// TwinCAT 3 PLC project Test
// ProgramVersion: 3.1.4026.26
// CompilerDefines: VISU_USEPROPERTYINFO
// libraries:
//   Tc2_Standard, * (Beckhoff Automation GmbH)
//   Tc2_System, * (Beckhoff Automation GmbH)
//   VisuDialogs, * (System)
//   VisuDialogs
// project tree:
//   DUTs/ Auto_Test_DB_DUT.TcDUT, Auto_Test_DUT.TcDUT, Barcode_Station_DUT.TcDUT, Charger_DUT.TcDUT, Gate_Station_DUT.TcDUT, Level_Keys_DUT.TcDUT, Profiling_Station_DUT.TcDUT, Shuttle_Position_UDT.TcDUT, U_DWORD_REAL1.TcDUT
//   DUTs/Carousel/ Chain_Control_DUT.TcDUT, Chain_Settings_DUT.TcDUT, E_Carousel_PopUpMotor.TcDUT, PopUp_Control_DUT.TcDUT, PopUp_Inputs_DUT.TcDUT, PopUp_Instruction_DUT.TcDUT, PopUp_Motors_DUT.TcDUT, PopUp_Motor_Settings_DUT.TcDUT, PopUp_Settings_DUT.TcDUT, PopUp_Side_Status_DUT.TcDUT, Roller_Control_DUT.TcDUT, Roller_Inputs_DUT.TcDUT, Roller_Instruction_DUT.TcDUT, Roller_Settings_DUT.TcDUT, TBCnv_Control_DUT.TcDUT, TBCnv_Settings_DUT.TcDUT, Turn_Table_Control_DUT.TcDUT, Turn_Table_Inputs_DUT.TcDUT, Turn_Table_Instruction_DUT.TcDUT, Turn_Table_Motor_DUT.TcDUT, Turn_Table_Settings_DUT.TcDUT
//   DUTs/Conveyors/ Buffer_Cnv_Control_DUT.TcDUT, Buffer_Cnv_Inputs_DUT.TcDUT, Buffer_Cnv_Settings_DUT.TcDUT, Cnv_Errors_DUT.TcDUT, Cnv_Inputs_DUT.TcDUT, Cnv_Instruction_DUT.TcDUT, Cnv_Interlock_DUT.TcDUT, Cnv_Level_Control_DUT.TcDUT, Cnv_Level_Inputs_DUT.TcDUT, Cnv_Level_Settings_DUT.TcDUT, Cnv_Motor_DUT.TcDUT, Cnv_Motor_Settings_DUT.TcDUT, Cnv_VTD_Control_DUT.TcDUT, Cnv_VTD_Settings_DUT.TcDUT, ECnv_Control_DUT.TcDUT, ECnv_Settings_DUT.TcDUT
//   DUTs/HMI/ ST_HMI_ConveyorCommand.TcDUT, ST_HMI_ConveyorStatus.TcDUT, ST_HMI_DeviceSummary.TcDUT, ST_HMI_GateCommand.TcDUT, ST_HMI_GateStatus.TcDUT, ST_HMI_GateSummary.TcDUT, ST_HMI_SystemCommand.TcDUT, ST_HMI_SystemStatus.TcDUT, ST_HMI_VtdCommand.TcDUT, ST_HMI_VtdOverview.TcDUT, ST_HMI_VtdStatus.TcDUT, ST_VTD_ManualHmiCommand.TcDUT, ST_VTD_ManualHmiStatus.TcDUT, ST_VTD_ManualSettings.TcDUT, ST_VTD_PdHmiCommand.TcDUT, ST_VTD_PdHmiStatus.TcDUT
//   DUTs/Safety_Stops/ Sfts_Control_DUT.TcDUT, Sfts_Inputs_DUT.TcDUT, Sfts_Instruction_DUT.TcDUT, Sfts_Settings_DUT.TcDUT
//   DUTs/SEW/ E_SEW_MovikitMode.TcDUT, ST_SEW_MovikitStatus.TcDUT, ST_SEW_ProcessInput5.TcDUT, ST_SEW_ProcessInput8.TcDUT, ST_SEW_VelocityScaling.TcDUT, ST_SEW_VelocityStatus.TcDUT
//   DUTs/System/ E_BarcodeState.TcDUT, ID_Decoded_DUT.TcDUT, OrderTable_DUT.TcDUT, System_DUT.TcDUT, System_Settings_DUT.TcDUT, WMS_OPC_UA_DUT.TcDUT
//   DUTs/VTD/ VTD_Control_DUT.TcDUT, VTD_Errors_DUT.TcDUT, VTD_Inputs_DUT.TcDUT, VTD_Instruction_DUT.TcDUT, VTD_Levels_DUT.TcDUT, VTD_Motor_DUT.TcDUT, VTD_Outputs_DUT.TcDUT, VTD_Settings_DUT.TcDUT, VTD_Shuttle_Interlock_DUT.TcDUT
//   / GlobalTextList.TcGTLO, PlcTask.TcTTO, TL_Test.TcTLO, Visualization Manager.TcVMO (not stored), VISU_TASK.TcTTO
//   GVLs/ Control.TcGVL, Errors.TcGVL, Settings.TcGVL, System.TcGVL, System_Control.TcGVL
//   GVLs/HMI/ CNV_HMI.TcGVL, CNV_HMI_IO.TcGVL, GVL_HMI_Carousel.TcGVL, GVL_HMI_CNV.TcGVL, GVL_HMI_Gates.TcGVL, GVL_HMI_System.TcGVL, GVL_HMI_VTD.TcGVL
//   GVLs/IO/ IO_Cards.TcGVL, IO_Chargers.TcGVL, IO_RemoteModules.TcGVL, IO_Safety.TcGVL, IO_VFDs.TcGVL
//   POUs/Conveyors/ Buffer_Conveyor_FB.TcPOU, FB_Conveyor_MotorInterlock.TcPOU
//   POUs/ DWORD_REAL.TcPOU, Inputs.TcPOU, MAIN.TcPOU, Outputs.TcPOU, Profile_Station_FC.TcPOU, Stack_Lights_FB.TcPOU
//   POUs/SEW/ FB_SEW_Drive.TcPOU, FB_SEW_ProcessDataTest.TcPOU, FB_SEW_VelocityDrive.TcPOU, FC_SEW_MovikitModeName.TcPOU, FC_VTD_PdHmiUpdateStatus.TcPOU
//   POUs/System/ Barcode_Station_FB.TcPOU, Conveyors_Transfer.TcPOU
//   POUs/System/Functions/ ByteArrayToString.TcPOU, FC_TIAParseDINT.TcPOU, FC_TIAScalarToken.TcPOU, FindBoolField.TcPOU, FindDINTFieldFragmented.TcPOU, FindIntField.TcPOU, FindINTFieldFragmented.TcPOU, FindStringField.TcPOU, ID_Decode_F.TcPOU, RemovePlusSign.TcPOU, Set_Bit_F.TcPOU
//   POUs/System/Tests/ FC_TestTIAFoundation.TcPOU, FC_TestTIAParsing.TcPOU
//   POUs/VTD/ FB_VTD_ManualControl.TcPOU, Light_Bars_FB.TcPOU, VTD_FB.TcPOU
//   VISUs/ Access_Gates.TcVIS, Alarms.TcVIS, Carrousel.TcVIS, CNV.TcVIS, CNV_Settings.TcVIS, Dialog.TcVIS, FP_Conveyor.TcVIS, FP_Drive.TcVIS, FP_Test.TcVIS, Header.TcVIS, ImagePool.TcIPO (not stored), Main.TcVIS, NavBar.TcVIS, Order_Table.TcVIS, Shuttles.TcVIS, teste.TcVIS, Visualization.TcVIS, VISU_Seeds.TcVIS, VTD.TcVIS, VTDManualTest.TcVIS, VTD_Settings.TcVIS
// real-time tasks:
//   TASK IoTask: cycle T#10ms, priority 1, ADS port 301
//   TASK PlcTask: cycle T#10ms, priority 20, ADS port 350
//   TASK VISU_TASK: cycle T#200000us, priority 30, ADS port 351
// I/O:
//   DEVICE Device 1 (EtherCAT), AmsNetId 10.1.179.234.2.1
//     Term 30 (EK1200) [EK1200-5000 EtherCAT Power supply (2A E-Bus)]
//       Term 3 (EL1809) [EL1809 16Ch. Dig. Input 24V, 3ms]
//       Term 4 (EL1809) [EL1809 16Ch. Dig. Input 24V, 3ms]
//       Term 5 (EL2809) [EL2809 16Ch. Dig. Output 24V, 0.5A]
//       Term 6 (EL2809) [EL2809 16Ch. Dig. Output 24V, 0.5A]
//       Term 7 (EL6910) [EL6910, TwinSAFE PLC]
//       Term 8 (EL1918) [EL1918, 8Ch. Safety Input 24V, TwinSAFE]
//         modules: Module 1 (FSOE), Module 2 (FSLOGIC)
//       Term 9 (EL2912) [EL2912, 2Ch. Safety Output 24V, 2A, TwinSAFE]
//         modules: Module 1 (FSOE), Module 2 (FSOUT), Module 3 (DEVICEIO), Module 4 (FSLOGIC)
//       Term 10 (EL9410) [EL9410 E-Bus Power Supplier  (Diagnostics)]
//       Term 11 (EK1322) [EK1322 2-port EtherCAT P junction with feed-in]
//       Term 12 (EK1322) [EK1322 2-port EtherCAT P junction with feed-in]
//       Term 13 (EK1322) [EK1322 2-port EtherCAT P junction with feed-in]
//         Box 14 (EPP2328-0002) [EPP2328-0002 4 CH. Dig. In, 3ms, 4 Ch. Dig. Out 24V, 2A, M12]
//       Term 43 (EL6633) [EL6633 PROFINET IO Controller]
//       Term 16 (EK1122) [EK1122 2 port EtherCAT junction]
//         Box 17 (CU1124) [CU1124 EtherCAT junction (4-ports)]
//         Box 19 (CU1128) [CU1128 6x EtherCAT junction]
//           Term 22 (CU1128-B) [CU1128 6x EtherCAT junction - Dev A]
//           Term 23 (CU1128-C) [CU1128 6x EtherCAT junction - Dev B]
//             Box 24 (MOVI-C Decentralized Electronics) [MOVI-C Decentralized Electronics]
//               modules: Module 1 (Standard 16 PD), Module 2 (Failsafe Container 28 Byte)
//             Box 25 (MOVI-C Decentralized Electronics) [MOVI-C Decentralized Electronics]
//               modules: Module 1 (Standard 16 PD), Module 2 (FSoE Safety IO 48 bit)
//             Box 45 (MOVI-C Decentralized Electronics) [MOVI-C Decentralized Electronics]
//               modules: Module 1 (Standard 16 PD), Module 2 (Failsafe Container 28 Byte)
//             Box 1 (MOVI-C MOVIPRO) [MOVI-C MOVIPRO]
//               modules: Module 1 (Standard 16 PD), Module 2 (FSoE Safety IO 48 bit)
//             Box 27 (MOVI-C Decentralized Electronics) [MOVI-C Decentralized Electronics]
//               modules: Module 1 (Standard 16 PD)
//             Box 47 (MOVI-C Decentralized Electronics) [MOVI-C Decentralized Electronics]
//               modules: Module 1 (Standard 16 PD)
//             Box 48 (MOVI-C Decentralized Electronics) [MOVI-C Decentralized Electronics]
//               modules: Module 1 (Standard 16 PD)
//             Box 49 (MOVI-C Decentralized Electronics) [MOVI-C Decentralized Electronics]
//               modules: Module 1 (Standard 16 PD)
//             Box 53 (MOVI-C Decentralized Electronics) [MOVI-C Decentralized Electronics]
//               modules: Module 1 (Standard 16 PD)
//   DEVICE Device 4 (COM Port)
// variable links:
//   Device 1 (EtherCAT) <-> Device 1 (EtherCAT)/Term 30 (EK1200)/Term 16 (EK1122)/Box 19 (CU1128)/Term 23 (CU1128-C)/Box 1 (MOVI-C MOVIPRO)
//     Term 30 (EK1200)/Term 7 (EL6910)/ConnectionInputs/Message_14 TxPDO <-> Module 2 (FSoE Safety IO 48 bit)/FSoE Safety Outputs 48 bit/FSOE
//     Term 30 (EK1200)/Term 7 (EL6910)/ConnectionOutputs/Message_14 RxPDO <-> Module 2 (FSoE Safety IO 48 bit)/FSoE Safety Inputs 48 bit/FSOE
//   Device 1 (EtherCAT) <-> Device 1 (EtherCAT)/Term 30 (EK1200)/Term 8 (EL1918)
//     Term 30 (EK1200)/Term 7 (EL6910)/ConnectionInputs/Message_13 TxPDO <-> Module 1 (FSOE)/FSoE Outputs/FSOE
//     Term 30 (EK1200)/Term 7 (EL6910)/ConnectionOutputs/Message_13 RxPDO <-> Module 1 (FSOE)/FSoE Inputs/FSOE
//   Test/Test Instance <-> Device 1 (EtherCAT)/Term 30 (EK1200)/Term 16 (EK1122)/Box 19 (CU1128)/Term 23 (CU1128-C)/Box 1 (MOVI-C MOVIPRO)
//     PlcTask Inputs/IO_VFDs.VTD_EcState <-> InfoData/State
//     PlcTask Inputs/IO_VFDs.VTD_PI_01 <-> Module 1 (Standard 16 PD)/Inputs 16 PD/PI 1
//     PlcTask Inputs/IO_VFDs.VTD_PI_02 <-> Module 1 (Standard 16 PD)/Inputs 16 PD/PI 2
//     PlcTask Inputs/IO_VFDs.VTD_PI_03 <-> Module 1 (Standard 16 PD)/Inputs 16 PD/PI 3
//     PlcTask Inputs/IO_VFDs.VTD_PI_04 <-> Module 1 (Standard 16 PD)/Inputs 16 PD/PI 4
//     PlcTask Inputs/IO_VFDs.VTD_PI_05 <-> Module 1 (Standard 16 PD)/Inputs 16 PD/PI 5
//     PlcTask Inputs/IO_VFDs.VTD_PI_06 <-> Module 1 (Standard 16 PD)/Inputs 16 PD/PI 6
//     PlcTask Inputs/IO_VFDs.VTD_PI_07 <-> Module 1 (Standard 16 PD)/Inputs 16 PD/PI 7
//     PlcTask Inputs/IO_VFDs.VTD_PI_08 <-> Module 1 (Standard 16 PD)/Inputs 16 PD/PI 8
//     PlcTask Inputs/IO_VFDs.VTD_WcState <-> WcState/WcState
//     PlcTask Outputs/IO_VFDs.VTD_PO_01 <-> Module 1 (Standard 16 PD)/Outputs 16 PD/PO 1
//     PlcTask Outputs/IO_VFDs.VTD_PO_02 <-> Module 1 (Standard 16 PD)/Outputs 16 PD/PO 2
//     PlcTask Outputs/IO_VFDs.VTD_PO_03 <-> Module 1 (Standard 16 PD)/Outputs 16 PD/PO 3
//     PlcTask Outputs/IO_VFDs.VTD_PO_04 <-> Module 1 (Standard 16 PD)/Outputs 16 PD/PO 4
//     PlcTask Outputs/IO_VFDs.VTD_PO_05 <-> Module 1 (Standard 16 PD)/Outputs 16 PD/PO 5
//     PlcTask Outputs/IO_VFDs.VTD_PO_06 <-> Module 1 (Standard 16 PD)/Outputs 16 PD/PO 6
//     PlcTask Outputs/IO_VFDs.VTD_PO_07 <-> Module 1 (Standard 16 PD)/Outputs 16 PD/PO 7
//     PlcTask Outputs/IO_VFDs.VTD_PO_08 <-> Module 1 (Standard 16 PD)/Outputs 16 PD/PO 8
//   Test/Test Instance <-> Device 1 (EtherCAT)/Term 30 (EK1200)/Term 7 (EL6910)
//     PlcTask Outputs/IO_Safety.ErrorAcknowledgement <-> StandardOutputs/Standard In Var 1
//     PlcTask Outputs/IO_Safety.Run <-> StandardOutputs/Standard In Var 2
//     PlcTask Outputs/IO_Safety.SEW_Safety_Reset <-> StandardOutputs/Standard In Var 10

CONFIGURATION Test
    RESOURCE PLC ON TwinCAT3
        TASK PlcTask(INTERVAL := T#10ms, PRIORITY := 20);
        TASK VISU_TASK(INTERVAL := T#200000us, PRIORITY := 30);
        PROGRAM MAIN WITH PlcTask : MAIN;
        PROGRAM VisuElems_Visu_Prg WITH VISU_TASK : VisuElems.Visu_Prg;
    END_RESOURCE
END_CONFIGURATION

// ---- DUTs/Auto_Test_DB_DUT.TcDUT
TYPE Auto_Test_DB_DUT :
STRUCT
	System: ARRAY[1..5] OF Auto_Test_DUT;
END_STRUCT
END_TYPE

// ---- DUTs/Auto_Test_DUT.TcDUT
TYPE Auto_Test_DUT :
STRUCT
	Duration:	TIME;
	Start_Time:	STRING[20];
	Stop_Time:	STRING[20];
	Time_Running:	TIME;
	Total_Duration:	TIME;
END_STRUCT
END_TYPE

// ---- DUTs/Barcode_Station_DUT.TcDUT
TYPE Barcode_Station_DUT :
STRUCT
	// Explicit capacity matches the default STRING length in the Siemens source.
	Start:	BOOL;
	Ready:	BOOL;
	Running:	BOOL;
	Done:	BOOL;
	Valid:	BOOL;
	Reading_Gate_number:	STRING(254);
	Reading_Gate_number_OLD:	STRING(254);
	Number_OF_Reading_Gates:	STRING(254);
	Number_OF_Reading_Gates_OLD:	STRING(254);
	Barcode:	STRING(254);
	Barcode_Old:	STRING(254);
END_STRUCT
END_TYPE

// ---- DUTs/Carousel/Chain_Control_DUT.TcDUT
// Internal state of the carousel chain conveyor (Control.Chain_Cnv).
// Same layout as ECnv_Control_DUT. Drive: SEW MOVIKIT Velocity Drive, 5 PD.
TYPE Chain_Control_DUT :
STRUCT
	Mode:	UINT;	// 0 Disabled, 1 Manual, 2 Semi-Auto, 3 Auto, 5 Maintenance
	Error:	BOOL;
	Warning:	UINT;
	Enabled:	BOOL;
	Stopped:	BOOL;
	Done:	BOOL;
	Running:	BOOL;
	Ready_For_Task:	BOOL;
	Current_Task_Type:	UINT;
	Current_Task_ID:	UINT;
	Cnv_Occupied:	BOOL;
	SM_State:	UINT;	// State machine value
	Motor:	Cnv_Motor_DUT;
	Instruction:	Cnv_Instruction_DUT;
	Inputs:	Cnv_Inputs_DUT;	// Forward/Backward_Sensor; VFD_* words not used with SEW
	Cnv_Errors:	Cnv_Errors_DUT;
END_STRUCT
END_TYPE

// ---- DUTs/Carousel/Chain_Settings_DUT.TcDUT
// Parameters of the carousel chain conveyor (Settings.Chain_Cnv). Based on ECnv_Settings_DUT.
// 0 = not configured: the function that uses the value is blocked.
TYPE Chain_Settings_DUT :
STRUCT
	ID:	DINT;	// XXYYZZ
	Motor:	Cnv_Motor_Settings_DUT;	// Same name as Control.<device>.Motor
END_STRUCT
END_TYPE

// ---- DUTs/Carousel/E_Carousel_PopUpMotor.TcDUT
// Motor of a carousel popup that is allowed to run (Control.Pop_Up_Cnv[n].Active_Motor).
// The values are the motor indices of the popup's FB_Conveyor_MotorInterlock instance.
{attribute 'qualified_only'}
TYPE E_Carousel_PopUpMotor :
(
    None := 0,          // No motor granted
    Lift := 1,          // Motors.Lift
    Transfer := 2       // Motors.Transfer
) INT;
END_TYPE

// ---- DUTs/Carousel/PopUp_Control_DUT.TcDUT
// Internal state of one carousel popup (Control.Pop_Up_Cnv[1..2]): lift + transfer conveyor.
// Based on Dallas PopUp_Cnv_Control; same header as ECnv_Control_DUT / Buffer_Cnv_Control_DUT.
// Motors.Lift and Motors.Transfer never run at the same time (Active_Motor, FB_Conveyor_MotorInterlock).
// Drives: SEW MOVIKIT Velocity Drive, 5 PD (Motor.stProcessInput / aProcessOutput in Cnv_Motor_DUT).
TYPE PopUp_Control_DUT :
STRUCT
	Mode:	UINT;	// 0 Disabled, 1 Manual, 2 Semi-Auto, 3 Auto, 5 Maintenance
	Error:	BOOL;
	Warning:	UINT;
	Enabled:	BOOL;
	Stopped:	BOOL;
	Done:	BOOL;
	Running:	BOOL;
	Ready_For_Task:	BOOL;
	Current_Task_Type:	UINT;
	Current_Task_ID:	UINT;
	Cnv_Occupied:	BOOL;
	SM_State:	UINT;	// State machine value
	Active_Side:	INT;	// Side 1..4 of the running transfer, 0 = none
	Inputs:	PopUp_Inputs_DUT;
	Side:	ARRAY[1..4] OF PopUp_Side_Status_DUT;	// 1/2 transfer Fwd/Rev end (Lift_Up), 3/4 Lift_Down level (pallet moved by the neighbour, e.g. Chain_Cnv)

	// Motor group: one motor at a time
	Motors:	PopUp_Motors_DUT;
	Active_Motor:	E_Carousel_PopUpMotor;	// Motor allowed to run, None = no motor granted
	Motor_Changeover:	BOOL;	// A motor is requested and waits until the other one stopped + Changeover_Time

	Instruction:	PopUp_Instruction_DUT;
	Cnv_Errors:	Cnv_Errors_DUT;
END_STRUCT
END_TYPE

// ---- DUTs/Carousel/PopUp_Inputs_DUT.TcDUT
// Sensors of one carousel popup (Control.Pop_Up_Cnv[n].Inputs). Written only by FC Inputs.
// Based on Dallas PopUp_Cnv_Inputs ("Lift Up" / "Lift Down") plus the popup pallet sensor.
// TRUE = condition present (invert NC sensors in FC Inputs).
TYPE PopUp_Inputs_DUT :
STRUCT
	Lift_Up:	BOOL;	// Lift at the top = transfer conveyor level
	Lift_Down:	BOOL;	// Lift at the bottom = chain level (pallet on Chain_Cnv, to confirm with the layout)
	Pallet_Present:	BOOL;	// Pallet on the popup (end of an inbound transfer)
END_STRUCT
END_TYPE

// ---- DUTs/Carousel/PopUp_Instruction_DUT.TcDUT
// Commands of one carousel popup (WMS / order table / HMI). Same members as Dallas PopUp_Cnv_Instruction.
TYPE PopUp_Instruction_DUT :
STRUCT
	Mode_Change:	UINT;	// Requested mode, see Mode
	Stop:	BOOL;
	Enable:	BOOL;
	Reset:	BOOL;
	Execute:	BOOL;	// Rising edge starts the task
	Task_ID:	UINT;
	Task_Metadata:	STRING;
	Transfer_To_ID:	DINT;	// Outbound: ID (XXYYZZ) of the receiving device
	Transfer_From_ID:	DINT;	// Inbound: ID (XXYYZZ) of the sending device
	Transfer_in_Progress:	BOOL;	// Written by the conveyor FB
	Inbound_Ready:	BOOL;	// Written by Conveyors_Transfer
	Transfer_Complete:	BOOL;
	Outbound_Ready:	BOOL;	// Written by Conveyors_Transfer
	Start_Transfer:	BOOL;
	Start_Transfer_Backward:	BOOL;	// Manual mode only

	// Manual mode
	Transfer_Fwd:	BOOL;	// Jog the transfer conveyor forward (only at Lift_Up)
	Transfer_Bwd:	BOOL;	// Jog the transfer conveyor backward (only at Lift_Up)
	Lift_Up:	BOOL;	// Auto: move the lift up. Manual: jog up
	Lift_Down:	BOOL;	// Auto: move the lift down. Manual: jog down
END_STRUCT
END_TYPE

// ---- DUTs/Carousel/PopUp_Motors_DUT.TcDUT
// Motors of one carousel popup (Control.Pop_Up_Cnv[n].Motors). They never run at the same time:
// PopUp_Conveyor_FB grants one motor at a time (FB_Conveyor_MotorInterlock, Active_Motor).
// Drives: SEW MOVIKIT Velocity Drive, 5 PD.
TYPE PopUp_Motors_DUT :
STRUCT
	Lift:	Cnv_Motor_DUT;	// Lift up / down (E_Carousel_PopUpMotor.Lift)
	Transfer:	Cnv_Motor_DUT;	// Transfer conveyor, runs only at Lift_Up (E_Carousel_PopUpMotor.Transfer)
END_STRUCT
END_TYPE

// ---- DUTs/Carousel/PopUp_Motor_Settings_DUT.TcDUT
// Motor parameters of one carousel popup (Settings.Pop_Up_Cnv[n].Motors).
// Same member names as PopUp_Motors_DUT in Control.
TYPE PopUp_Motor_Settings_DUT :
STRUCT
	Lift:	Cnv_Motor_Settings_DUT;	// Transfer_Time = lift travel watchdog
	Transfer:	Cnv_Motor_Settings_DUT;
END_STRUCT
END_TYPE

// ---- DUTs/Carousel/PopUp_Settings_DUT.TcDUT
// Parameters of one carousel popup (Settings.Pop_Up_Cnv[1..2]). Based on Dallas PopUp_Cnv_Settings;
// the G120 hardware IDs are replaced by the SEW scaling of each drive (Motors.<motor>.Drive).
// 0 = not configured: the function that uses the value is blocked.
TYPE PopUp_Settings_DUT :
STRUCT
	ID:	DINT;	// XXYYZZ
	Side_ID:	ARRAY[1..4] OF DINT;	// Neighbour ID per side, 0 = none. 1/2 transfer Fwd/Rev end (Lift_Up), 3/4 Lift_Down level
	Side_Boost_Time:	ARRAY[1..4] OF UINT;	// [s] start boost per side, 0 = none (Dallas TimeStartBoost_PxToPy)
	Boost_Speed:	UINT := 100;	// Units of Motors.Transfer.Speed

	// Motor group: Lift and Transfer never run at the same time
	Motors:	PopUp_Motor_Settings_DUT;
	Changeover_Time:	UINT;	// [ms] all motors stopped before the other motor may start (brake closed), 0 = not configured
END_STRUCT
END_TYPE

// ---- DUTs/Carousel/PopUp_Side_Status_DUT.TcDUT
// Device on one side of a popup (Control.Pop_Up_Cnv[n].Side[1..4]). Written every cycle by Conveyors_Transfer.
// Replaces the hard-coded neighbour reads of the Dallas PConveyor FBs.
TYPE PopUp_Side_Status_DUT :
STRUCT
	In_Position:	BOOL;	// Neighbour aligned with the popup (VTD at the level, turntable at the station). TRUE for fixed conveyors
	Inbound_Ready:	BOOL;	// Neighbour can receive a pallet
	Running:	BOOL;	// Neighbour transport motor turning (handshake before sending)
	Occupied:	BOOL;	// Neighbour detects the pallet (end of an outbound transfer)
END_STRUCT
END_TYPE

// ---- DUTs/Carousel/Roller_Control_DUT.TcDUT
// Internal state of one carousel roller conveyor (Control.Roller_Cnv[1..5]).
// Same layout as ECnv_Control_DUT. Drive: SEW MOVIKIT Velocity Drive, 5 PD.
TYPE Roller_Control_DUT :
STRUCT
	Mode:	UINT;	// 0 Disabled, 1 Manual, 2 Semi-Auto, 3 Auto, 5 Maintenance
	Error:	BOOL;
	Warning:	UINT;
	Enabled:	BOOL;
	Stopped:	BOOL;
	Done:	BOOL;
	Running:	BOOL;
	Ready_For_Task:	BOOL;
	Current_Task_Type:	UINT;
	Current_Task_ID:	UINT;
	Cnv_Occupied:	BOOL;
	SM_State:	UINT;	// State machine value
	Motor:	Cnv_Motor_DUT;
	Instruction:	Roller_Instruction_DUT;
	Inputs:	Roller_Inputs_DUT;
	Cnv_Errors:	Cnv_Errors_DUT;
END_STRUCT
END_TYPE

// ---- DUTs/Carousel/Roller_Inputs_DUT.TcDUT
// Sensors of one carousel roller conveyor (Control.Roller_Cnv[n].Inputs). Written only by FC Inputs.
// Based on Cnv_Inputs_DUT and Dallas Inbound/Outbound_Cnv_Inputs. The VFD_* words are not needed:
// with SEW the drive data is in Motor.stProcessInput. TRUE = condition present (invert NC sensors in FC Inputs).
TYPE Roller_Inputs_DUT :
STRUCT
	Forward_Sensor:	BOOL;	// Pallet at the forward end
	Backward_Sensor:	BOOL;	// Pallet at the backward end
	Fork_Lift_Detect:	BOOL;	// Forklift in the station (forklift stations only, FALSE otherwise)
END_STRUCT
END_TYPE

// ---- DUTs/Carousel/Roller_Instruction_DUT.TcDUT
// Commands of one carousel roller conveyor. Cnv_Instruction_DUT + Dallas InCnv/OutCnv_Instruction station flags.
TYPE Roller_Instruction_DUT :
STRUCT
	Mode_Change:	UINT;	// Requested mode, see Mode
	Stop:	BOOL;
	Enable:	BOOL;
	Reset:	BOOL;
	Execute:	BOOL;	// Rising edge starts the task
	Task_ID:	UINT;
	Task_Metadata:	STRING;
	Transfer_To_ID:	DINT;	// Outbound: ID (XXYYZZ) of the receiving device
	Transfer_From_ID:	DINT;	// Inbound: ID (XXYYZZ) of the sending device
	Transfer_in_Progress:	BOOL;	// Written by the conveyor FB
	Inbound_Ready:	BOOL;	// Written by Conveyors_Transfer
	Transfer_Complete:	BOOL;
	Outbound_Ready:	BOOL;	// Written by Conveyors_Transfer
	Start_Transfer:	BOOL;
	Start_Transfer_Backward:	BOOL;	// Manual mode only
	Foward:	BOOL;	// Manual jog forward (spelling as Cnv_Instruction_DUT)
	Backward:	BOOL;	// Manual jog backward

	// Forklift stations (Dallas InConveyor_FB / OutConveyor_FB)
	Automatic_Start:	BOOL;	// PLC -> WMS: pallet placed, no forklift for No_Forklift_Detect_Timer
	Empty:	BOOL;	// PLC -> WMS: station empty, no forklift for No_Forklift_Detect_Timer
END_STRUCT
END_TYPE

// ---- DUTs/Carousel/Roller_Settings_DUT.TcDUT
// Parameters of one carousel roller conveyor (Settings.Roller_Cnv[1..5]).
// Based on ECnv_Settings_DUT / Buffer_Cnv_Settings_DUT and Dallas Inbound/Outbound_Cnv_Settings.
// 0 = not configured: the function that uses the value is blocked.
TYPE Roller_Settings_DUT :
STRUCT
	ID:	DINT;	// XXYYZZ
	Barcode_ID:	UINT;	// Barcode station at this roller, 0 = none
	Motor:	Cnv_Motor_Settings_DUT;	// Same name as Control.<device>.Motor
	No_Forklift_Detect_Timer:	UINT;	// [s] forklift stations: time without forklift before Automatic_Start / Empty
END_STRUCT
END_TYPE

// ---- DUTs/Carousel/TBCnv_Control_DUT.TcDUT
// Internal state of the turntable roller conveyor (Control.TBCnv).
// Same layout as ECnv_Control_DUT. Drive: SEW MOVIKIT Velocity Drive, 5 PD.
TYPE TBCnv_Control_DUT :
STRUCT
	Mode:	UINT;	// 0 Disabled, 1 Manual, 2 Semi-Auto, 3 Auto, 5 Maintenance
	Error:	BOOL;
	Warning:	UINT;
	Enabled:	BOOL;
	Stopped:	BOOL;
	Done:	BOOL;
	Running:	BOOL;
	Ready_For_Task:	BOOL;
	Current_Task_Type:	UINT;
	Current_Task_ID:	UINT;
	Cnv_Occupied:	BOOL;
	SM_State:	UINT;	// State machine value
	Motor:	Cnv_Motor_DUT;
	Instruction:	Cnv_Instruction_DUT;
	Inputs:	Cnv_Inputs_DUT;	// Forward/Backward_Sensor; VFD_* words not used with SEW
	Cnv_Errors:	Cnv_Errors_DUT;

	// Interlock with Control.Turn_Table: turntable rotation and turntable roller never run at the same time
	Interlock:	Cnv_Interlock_DUT;	// Run_Request / Motor_Stopped by this FB, Run_Allowed by the group FB_Conveyor_MotorInterlock
END_STRUCT
END_TYPE

// ---- DUTs/Carousel/TBCnv_Settings_DUT.TcDUT
// Parameters of the turntable roller conveyor (Settings.TBCnv). Based on ECnv_Settings_DUT.
// 0 = not configured: the function that uses the value is blocked.
TYPE TBCnv_Settings_DUT :
STRUCT
	ID:	DINT;	// XXYYZZ
	Motor:	Cnv_Motor_Settings_DUT;	// Same name as Control.<device>.Motor
END_STRUCT
END_TYPE

// ---- DUTs/Carousel/Turn_Table_Control_DUT.TcDUT
// Internal state of the turntable (Control.Turn_Table): rotation axis only, the conveyor on it is Control.TBCnv.
// Same header as the conveyor DUTs. Drive: SEW MOVIKIT Positioning Drive (8 PD).
TYPE Turn_Table_Control_DUT :
STRUCT
	Mode:	UINT;	// 0 Disabled, 1 Manual, 2 Semi-Auto, 3 Auto, 5 Maintenance
	Error:	BOOL;
	Warning:	UINT;
	Enabled:	BOOL;
	Stopped:	BOOL;
	Done:	BOOL;
	Running:	BOOL;
	Ready_For_Task:	BOOL;
	Current_Task_Type:	UINT;
	Current_Task_ID:	UINT;
	SM_State:	UINT;	// State machine value
	Current_Position:	UINT;	// Station 1..4 reached, 0 = between stations / unknown
	In_Position:	BOOL;	// At Current_Position within Settings.Turn_Table.Position_Tolerance
	Motor:	Turn_Table_Motor_DUT;
	Instruction:	Turn_Table_Instruction_DUT;
	Inputs:	Turn_Table_Inputs_DUT;
	Cnv_Errors:	Cnv_Errors_DUT;

	// Interlock with Control.TBCnv: turntable rotation and turntable roller never run at the same time
	Interlock:	Cnv_Interlock_DUT;	// Run_Request / Motor_Stopped by this FB, Run_Allowed by the group FB_Conveyor_MotorInterlock
END_STRUCT
END_TYPE

// ---- DUTs/Carousel/Turn_Table_Inputs_DUT.TcDUT
// Sensors of the turntable (Control.Turn_Table.Inputs). Written only by FC Inputs.
// Encoder: SSI on the remote module "ENCODER (EPP5001-0002)" (candidate, AGENTS.md "Turntable").
// Bit length, Gray/binary code, resolution, direction and status bits are NOT confirmed:
// keep the values raw and never forward an invalid position to the drive.
TYPE Turn_Table_Inputs_DUT :
STRUCT
	Encoder_Value_Raw:	UDINT;	// EPP5001 SSI value, raw (format to confirm)
	Encoder_Status_Raw:	WORD;	// EPP5001 status, raw (width and bits to confirm)
	Encoder_WcState_Error:	BOOL;	// WcState of the encoder module (TRUE = data invalid)
	Encoder_EcState:	UINT;	// InfoData.State of the encoder module (8 = OP)
END_STRUCT
END_TYPE

// ---- DUTs/Carousel/Turn_Table_Instruction_DUT.TcDUT
// Commands of the turntable. Same first fields as Cnv_Instruction_DUT.
TYPE Turn_Table_Instruction_DUT :
STRUCT
	Mode_Change:	UINT;	// Requested mode, see Mode
	Stop:	BOOL;
	Enable:	BOOL;
	Reset:	BOOL;
	Execute:	BOOL;	// Rising edge starts the task
	Task_ID:	UINT;
	Task_Metadata:	STRING;
	Target_Position:	UINT;	// Station 1..4 to rotate to (Settings.Turn_Table.Position[n]), 0 = none
	Start_Rotation:	BOOL;
	Rotation_in_Progress:	BOOL;	// Written by the turntable FB

	// Manual mode
	Rotate_CW:	BOOL;	// Jog clockwise
	Rotate_CCW:	BOOL;	// Jog counter-clockwise
END_STRUCT
END_TYPE

// ---- DUTs/Carousel/Turn_Table_Motor_DUT.TcDUT
// Turntable drive: SEW MOVI-C with MOVIKIT Positioning Drive, 8 PD (confirm in MOVISUITE, AGENTS.md).
// Same layout as VTD_Motor_DUT. Raw process data is filled by FC Inputs and sent by FC Outputs.
TYPE Turn_Table_Motor_DUT :
STRUCT
	stProcessInput:	ST_SEW_ProcessInput8;	// PI 1..8 + EtherCAT diagnostics, written by Inputs
	aProcessOutput:	ARRAY[1..8] OF UINT;	// PO 1..8 raw, read by Outputs
	stStatus:	ST_SEW_MovikitStatus;	// Decoded drive status, written by the turntable FB
END_STRUCT
END_TYPE

// ---- DUTs/Carousel/Turn_Table_Settings_DUT.TcDUT
// Parameters of the turntable (Settings.Turn_Table). Number of stations to confirm (Rev 9).
// 0 = not configured: the function that uses the value is blocked.
TYPE Turn_Table_Settings_DUT :
STRUCT
	ID:	DINT;	// XXYYZZ
	Rotation_Time:	UINT;	// [s] rotation watchdog
	Full_Speed:	UINT;	// [%] automatic rotation
	Manual_Speed:	UINT;	// [%] manual jog

	// Station positions, drive user units (MOVIKIT Positioning). 0 = not taught: rotation to that station blocked
	Position:	ARRAY[1..4] OF DINT;
	Position_Tolerance:	DINT;	// [user units] in-position window

	// Interlock with the turntable roller conveyor (Control.TBCnv)
	Changeover_Time:	UINT;	// [ms] rotation and roller both stopped before the other may start, 0 = not configured

	// SEW MOVIKIT scaling (user units from MOVISUITE), as VTD_Settings_DUT
	SEW_Speed_At_100pct:	INT;	// PO 2 speed setpoint [user units] for 100 %
	SEW_Ramp_At_100pct:	UINT;	// PO 3/PO 4 acceleration/deceleration [user units] for 100 %
END_STRUCT
END_TYPE

// ---- DUTs/Charger_DUT.TcDUT
TYPE Charger_DUT :
STRUCT
	Output_Voltage:	REAL;                   	//Actual Output Voltage  
	Output_Current:	REAL;                       //Actual Output Current  
	Set_Voltage_Feedback:	REAL;               //Set Voltage Value      
	Set_Current_Feedback:	REAL;               //Set Current Value      
	Charging_Start:	BOOL;                       //Charging Running Status
	Set_Voltage_Output:	REAL;                   //Issue Target Voltage   
	Set_Current_Output:	REAL;                   //Issue Target Current   
	Start_Charging:	BOOL;                       //Start Charging Command 
	Stop_Charging:	BOOL;                       //Stop Charging Command  
	Confirm_Voltage_Current_Setting:	BOOL;   //Confirmation Command   
END_STRUCT
END_TYPE

// ---- DUTs/Conveyors/Buffer_Cnv_Control_DUT.TcDUT
TYPE Buffer_Cnv_Control_DUT :
STRUCT
	Mode:	UINT;
	Error:	BOOL;
	Warning:	UINT;
	Enabled:	BOOL;
	Stopped:	BOOL;
	Done:	BOOL;
	Running:	BOOL;
	Ready_For_Task:	BOOL;
	Current_Task_Type:	UINT;
	Current_Task_ID:	UINT;
	Cnv_Occupied:	BOOL;
	SM_State:	UINT;
	Motor:	Cnv_Motor_DUT;
	Instruction:	Cnv_Instruction_DUT;
	Inputs:	Buffer_Cnv_Inputs_DUT;
	Safety_Stop_Cnrl:	Sfts_Control_DUT;
	Cnv_Errors:	Cnv_Errors_DUT;
END_STRUCT
END_TYPE

// ---- DUTs/Conveyors/Buffer_Cnv_Inputs_DUT.TcDUT
TYPE Buffer_Cnv_Inputs_DUT :
STRUCT
	Forward_Sensor:	BOOL;
	Backward_Sensor:	BOOL;
	Shuttle_High:	BOOL;
	VFD_Status:	WORD;
	VFD_Speed_Actual:	INT;
	VFD_ActualCurrent:	INT;
	VFD_ActualTorque:	INT;
END_STRUCT
END_TYPE

// ---- DUTs/Conveyors/Buffer_Cnv_Settings_DUT.TcDUT
TYPE Buffer_Cnv_Settings_DUT :
STRUCT
	ID:	DINT;
	Barcode_ID:	UINT;
	Cnv_Level:	UINT;
	TC_Time:	UINT;
	Transfer_Time:	UINT;
	Pallet_Align_Time:	UINT;
	Slow_Speed:	UINT;
	Full_Speed:	UINT;
	Manual_Speed:	UINT;
	Safety_stop_Timeout:	UINT;

	// SEW MOVIKIT Velocity scaling (user units from MOVISUITE). 0 = not configured: the conveyor does not move.
	// Motor.Speed uses the units of Full_Speed / Slow_Speed / Manual_Speed.
	// Legacy Siemens scaling for reference: Motor.Speed 130 = 1865 rpm (G120 reference speed).
	rSewSpeedPerUnit:	REAL;     // PO 2 setpoint [user units] per 1 unit of Motor.Speed
	uiSewAcceleration:	UINT;    // PO 3 acceleration [user units]
	uiSewDeceleration:	UINT;    // PO 4 deceleration [user units]
END_STRUCT
END_TYPE

// ---- DUTs/Conveyors/Cnv_Errors_DUT.TcDUT
TYPE Cnv_Errors_DUT :
STRUCT
	// Bit fields. WORD (was UINT, as in the Siemens source) so that the words can be
	// passed to Set_Bit_F, whose VAR_IN_OUT Variavel is a WORD.
	Error_Word_1:	WORD;
	Error_Word_2:	WORD;
	Error_Word_3:	WORD;
	Error_Word_4:	WORD;
END_STRUCT
END_TYPE

// ---- DUTs/Conveyors/Cnv_Inputs_DUT.TcDUT
TYPE Cnv_Inputs_DUT :
STRUCT
	Forward_Sensor:	BOOL;
	Backward_Sensor:	BOOL;
	VFD_Status:	WORD;
	VFD_Speed_Actual:	INT;
	VFD_ActualCurrent:	INT;
	VFD_ActualTorque:	INT;
END_STRUCT
END_TYPE

// ---- DUTs/Conveyors/Cnv_Instruction_DUT.TcDUT
TYPE Cnv_Instruction_DUT :
STRUCT
	Mode_Change:	UINT;
	Stop:	BOOL;
	Enable:	BOOL;
	Reset:	BOOL;
	Execute:	BOOL;
	Task_ID:	UINT;
	Task_Metadata:	STRING;
	Transfer_To_ID:	DINT;
	Transfer_From_ID:	DINT;
	Transfer_in_Progress:	BOOL;
	Inbound_Ready:	BOOL;
	Transfer_Complete:	BOOL;
	Outbound_Ready:	BOOL;
	Start_Transfer:	BOOL;
	Foward:	BOOL;
	Backward:	BOOL;
END_STRUCT
END_TYPE

// ---- DUTs/Conveyors/Cnv_Interlock_DUT.TcDUT
// Motor interlock between two or more devices whose motors must not run at the same time
// (for example Control.Turn_Table rotation and Control.TBCnv roller).
// One FB_Conveyor_MotorInterlock instance per group grants one motor at a time.
// Functional interlock in the standard PLC, NOT a safety function.
TYPE Cnv_Interlock_DUT :
STRUCT
	Run_Request:	BOOL;	// Device FB -> interlock: the device wants to run its motor
	Motor_Stopped:	BOOL;	// Device FB -> interlock: motor not turning and output stage off
	Run_Allowed:	BOOL;	// Interlock -> device FB: the motor may run. FALSE = stop and do not start
END_STRUCT
END_TYPE

// ---- DUTs/Conveyors/Cnv_Level_Control_DUT.TcDUT
TYPE Cnv_Level_Control_DUT :
STRUCT
	Cnv1:	Buffer_Cnv_Control_DUT;
	Cnv2:	Buffer_Cnv_Control_DUT;
END_STRUCT
END_TYPE

// ---- DUTs/Conveyors/Cnv_Level_Inputs_DUT.TcDUT
TYPE Cnv_Level_Inputs_DUT :
STRUCT
	Cnv1_Inputs:	Buffer_Cnv_Inputs_DUT;
	Cnv2_Inputs:	Buffer_Cnv_Inputs_DUT;
END_STRUCT
END_TYPE

// ---- DUTs/Conveyors/Cnv_Level_Settings_DUT.TcDUT
TYPE Cnv_Level_Settings_DUT :
STRUCT
	Cnv1:	Buffer_Cnv_Settings_DUT;
	Cnv2:	Buffer_Cnv_Settings_DUT;
END_STRUCT
END_TYPE

// ---- DUTs/Conveyors/Cnv_Motor_DUT.TcDUT
TYPE Cnv_Motor_DUT :
STRUCT
	Enable:	BOOL;
	Enabled:	BOOL;
	Ready:	BOOL;
	Forward:	BOOL;
	Reverse:	BOOL;
	Speed:	REAL;
	Speed_Actual:	REAL;
	Actual_Current:	REAL;
	Actual_Torque:	UINT;
	Config_Axis:	WORD;
	Error:	BOOL;
	Status:	WORD;
	Communication_Error:	WORD;
	Lockout:	BOOL;

	// SEW MOVIKIT Velocity Drive, "5 PD" profile (buffer and roller conveyors).
	// stProcessInput is written only by FC Inputs; aProcessOutput is read only by FC Outputs.
	stProcessInput:	ST_SEW_ProcessInput5;   // PI 1..5 + EtherCAT diagnostics, written by Inputs
	aProcessOutput:	ARRAY[1..5] OF UINT;    // PO 1..5 raw, written by the conveyor FB, read by Outputs
	stStatus:	ST_SEW_VelocityStatus;          // Decoded drive status, written by the conveyor FB
END_STRUCT
END_TYPE

// ---- DUTs/Conveyors/Cnv_Motor_Settings_DUT.TcDUT
// Parameters of one conveyor motor (SEW MOVIKIT Velocity Drive, 5 PD).
// Settings counterpart of Cnv_Motor_DUT: Settings.<Device>.Motor(s) mirrors Control.<Device>.Motor(s).
// Speeds use the units of Cnv_Motor_DUT.Speed (Dallas: % of the drive range).
// 0 = not configured: the function that uses the value is blocked.
TYPE Cnv_Motor_Settings_DUT :
STRUCT
	TC_Time:	UINT;
	Transfer_Time:	UINT;	// [s] watchdog of a transfer (or of a lift travel)
	Slow_Speed:	UINT;	// Units of Motor.Speed
	Full_Speed:	UINT;	// Units of Motor.Speed
	Manual_Speed:	UINT;	// Units of Motor.Speed
	Drive:	ST_SEW_VelocityScaling;	// SEW MOVIKIT Velocity scaling and ramps
END_STRUCT
END_TYPE

// ---- DUTs/Conveyors/Cnv_VTD_Control_DUT.TcDUT
TYPE Cnv_VTD_Control_DUT :
STRUCT
	Cnv_Level:	ARRAY[1..6] OF Cnv_Level_Control_DUT;
END_STRUCT
END_TYPE

// ---- DUTs/Conveyors/Cnv_VTD_Settings_DUT.TcDUT
TYPE Cnv_VTD_Settings_DUT :
STRUCT
	Cnv_Level:	ARRAY[2..6] OF Cnv_Level_Settings_DUT;
END_STRUCT
END_TYPE

// ---- DUTs/Conveyors/ECnv_Control_DUT.TcDUT
TYPE ECnv_Control_DUT :
STRUCT
	Mode:	UINT;
	Error:	BOOL;
	Warning:	UINT;
	Enabled:	BOOL;
	Stopped:	BOOL;
	Done:	BOOL;
	Running:	BOOL;
	Ready_For_Task:	BOOL;
	Current_Task_Type:	UINT;
	Current_Task_ID:	UINT;
	Cnv_Occupied:	BOOL;
	SM_State:	UINT;
	Motor:	Cnv_Motor_DUT;
	Instruction:	Cnv_Instruction_DUT;
	Inputs:	Cnv_Inputs_DUT;
	Cnv_Errors:	Cnv_Errors_DUT;
END_STRUCT
END_TYPE

// ---- DUTs/Conveyors/ECnv_Settings_DUT.TcDUT
TYPE ECnv_Settings_DUT :
STRUCT
	ID:	DINT;
	Barcode_ID:	UINT;
	Cnv_Level:	UINT;
	TC_Time:	UINT;
	Transfer_Time:	UINT;
	Pallet_Align_Time:	UINT;
	Slow_Speed:	UINT;
	Full_Speed:	UINT;
	Manual_Speed:	UINT;
END_STRUCT
END_TYPE

// ---- DUTs/Gate_Station_DUT.TcDUT
TYPE Gate_Station_DUT :
STRUCT
	Requested_Access:	BOOL;
	Secure_Access:	BOOL;
	Safe_To_Restart:	BOOL;
END_STRUCT
END_TYPE

// ---- DUTs/HMI/ST_HMI_ConveyorCommand.TcDUT
// HMI -> PLC: commands for the device selected on the screens CNV / Carrousel.
// All Tap buttons. Jog, lift and rotate are hold-to-run (TRUE while pressed).
TYPE ST_HMI_ConveyorCommand :
STRUCT
    bModeManual : BOOL;
    bModeSemi : BOOL;
    bModeAuto : BOOL;
    bEnable : BOOL;
    bStop : BOOL;
    bReset : BOOL;
    bJogForward : BOOL;
    bJogBackward : BOOL;
    bLiftUp : BOOL;
    bLiftDown : BOOL;
    bRotateCw : BOOL;
    bRotateCcw : BOOL;
END_STRUCT
END_TYPE

// ---- DUTs/HMI/ST_HMI_ConveyorStatus.TcDUT
// PLC -> HMI: status of one conveyor-type device (extractor, buffer level, popup,
// roller, chain, turntable) for the screens CNV and Carrousel.
TYPE ST_HMI_ConveyorStatus :
STRUCT
    sName : STRING(20);            // For example 'Buffer L1', 'PopUp 2'
    bSelected : BOOL;              // Shown in the detail panel
    bEnabled : BOOL;
    bError : BOOL;
    bWarning : BOOL;
    bStopped : BOOL;
    bRunning : BOOL;
    bReadyForTask : BOOL;
    bOccupied : BOOL;
    bModeManual : BOOL;
    bModeSemi : BOOL;
    bModeAuto : BOOL;
    bForwardSensor : BOOL;
    bBackwardSensor : BOOL;
    bShuttleHigh : BOOL;           // Buffers only
    sMotorDirection : STRING(12);  // 'Stopped', 'Forward', 'Backward'
    iSpeedRequested_pct : INT;
    iSpeedActual_pct : INT;
    rCurrent_A : REAL;
    rTorque_pct : REAL;
    diTransferToId : DINT;
    diTransferFromId : DINT;
    uiStateMachine : UINT;
    bHasLift : BOOL;               // Popups
    bLiftUp : BOOL;
    bLiftDown : BOOL;
    bHasRotation : BOOL;           // Turntable
    rAngle_deg : REAL;
END_STRUCT
END_TYPE

// ---- DUTs/HMI/ST_HMI_DeviceSummary.TcDUT
// PLC -> HMI: summary of one device (conveyor, popup, roller, chain, turntable)
// for the tiles of the screen Main.
TYPE ST_HMI_DeviceSummary :
STRUCT
    bEnabled : BOOL;        // Device / drive enabled
    bRunning : BOOL;        // Moving (motor turning)
    bOccupied : BOOL;       // Pallet present
    bError : BOOL;          // Fault active (tile turns red)
    bWarning : BOOL;        // Warning active
    bManualMode : BOOL;     // Device in manual mode
    uiStateMachine : UINT;  // Current state number, diagnostics only
END_STRUCT
END_TYPE

// ---- DUTs/HMI/ST_HMI_GateCommand.TcDUT
// HMI -> PLC: gate requests (Tap). A request only; unlocking stays with the safety logic.
TYPE ST_HMI_GateCommand :
STRUCT
    bRequestAccess : BOOL;
    bReset : BOOL;
END_STRUCT
END_TYPE

// ---- DUTs/HMI/ST_HMI_GateStatus.TcDUT
// PLC -> HMI: status of one access gate for the screen Access_Gates (display only).
TYPE ST_HMI_GateStatus :
STRUCT
    bClosed : BOOL;
    bLocked : BOOL;
    bAccessRequested : BOOL;
    bAccessGranted : BOOL;    // Gate_Station.Secure_Access
    bSafeToRestart : BOOL;    // Gate_Station.Safe_To_Restart
    bError : BOOL;
END_STRUCT
END_TYPE

// ---- DUTs/HMI/ST_HMI_GateSummary.TcDUT
// PLC -> HMI: access gate summary for the screen Main (display only, not a safety function).
TYPE ST_HMI_GateSummary :
STRUCT
    bClosed : BOOL;          // Door closed
    bLocked : BOOL;          // Door locked
    bAccessRequested : BOOL; // Operator requested access
    bError : BOOL;           // Fault active (tile turns red)
END_STRUCT
END_TYPE

// ---- DUTs/HMI/ST_HMI_SystemCommand.TcDUT
// HMI -> PLC: commands of the screen Main.
TYPE ST_HMI_SystemCommand :
STRUCT
    bResetAll : BOOL;  // Tap - reset of all devices of this system (evaluated on the rising edge)
    bSafetyReset : BOOL;  // Tap - safety reset request (rising edge in MAIN -> one 500 ms pulse on IO_Safety.ErrorAcknowledgement
                          // and IO_Safety.SEW_Safety_Reset). The TwinSAFE logic decides whether the reset is accepted.
END_STRUCT
END_TYPE

// ---- DUTs/HMI/ST_HMI_SystemStatus.TcDUT
// PLC -> HMI: status of this system (one VTD panel) for the header and the screen Main.
TYPE ST_HMI_SystemStatus :
STRUCT
    iSystemNumber : INT;       // VTD number of this panel (1..10)
    sSystemName : STRING(40);  // For example 'VTD 1'
    dtNow : DT;                // PLC local time shown in the header
    bAutoMode : BOOL;
    bManualMode : BOOL;
    bSafetyOk : BOOL;          // Safety circuit OK (TwinSAFE status, display only)
    bSafetyResetActive : BOOL; // Safety reset pulse active (written by MAIN)
    bError : BOOL;
    bWarning : BOOL;
    uiActiveAlarms : UINT;
    sMessage : STRING(80);     // Operator message line
    bMessageAlarm : BOOL;      // TRUE = message line red
END_STRUCT
END_TYPE

// ---- DUTs/HMI/ST_HMI_VtdCommand.TcDUT
// HMI -> PLC: commands of the screen VTD (all Tap buttons, evaluated on the rising edge).
TYPE ST_HMI_VtdCommand :
STRUCT
    bModeManual : BOOL;
    bModeSemi : BOOL;
    bModeAuto : BOOL;
    bStop : BOOL;
    bReset : BOOL;
END_STRUCT
END_TYPE

// ---- DUTs/HMI/ST_HMI_VtdOverview.TcDUT
// PLC -> HMI: VTD summary for the screen Main.
TYPE ST_HMI_VtdOverview :
STRUCT
    stSummary : ST_HMI_DeviceSummary;
    uiCurrentLevel : UINT;  // 0 = between levels
    uiTargetLevel : UINT;   // 0 = no target
    rPosition_mm : REAL;    // Carriage position in mm (only after the MOVISUITE user units are confirmed)
    bDocked : BOOL;
    bPalletLoaded : BOOL;
    bShuttleLoaded : BOOL;
END_STRUCT
END_TYPE

// ---- DUTs/HMI/ST_HMI_VtdStatus.TcDUT
// PLC -> HMI: status of the VTD for the screen VTD.
TYPE ST_HMI_VtdStatus :
STRUCT
    // State
    bEnabled : BOOL;
    bError : BOOL;
    bStopped : BOOL;
    bRunning : BOOL;
    bDocked : BOOL;
    bSafetyOk : BOOL;                  // Display only
    bModeManual : BOOL;
    bModeSemi : BOOL;
    bModeAuto : BOOL;
    sPalletType : STRING(20);
    uiCurrentLevel : UINT;             // 0 = between levels
    uiLevelBelow : UINT;
    uiStateMachine : UINT;
    sDockingPinState : STRING(20);     // 'Extended', 'Retracted', ...
    sBarcode : STRING(40);

    // Position and drive
    rLePosition_mm : REAL;             // DL50 position
    rLeSpeed_mm_s : REAL;
    diAbsoluteEncoder : DINT;
    iEncoderDelta : INT;
    bLinearEncoderError : BOOL;
    bAbsoluteEncoderError : BOOL;
    bBarcodeError : BOOL;
    iSetpoint_pct : INT;
    iVelocity_pct : INT;
    rVelocity_mm_s : REAL;
    rCurrent_A : REAL;
    iTorque_pct : INT;
    bMotorReady : BOOL;

    // Levels and limit switches
    abLevelReached : ARRAY[1..8] OF BOOL;
    arLevelPosition_mm : ARRAY[1..8] OF REAL;  // Teach values
    bUpperOvertravel : BOOL;
    bUpperLimit : BOOL;
    bLowerLimit : BOOL;
    bLowerOvertravel : BOOL;

    // Signals
    bLevelDetect1 : BOOL;
    bLevelDetect2 : BOOL;
    bUltimateSlowdown : BOOL;
    bUltimateCreep : BOOL;
    bDp1Extended : BOOL;
    bDp2Extended : BOOL;
    bDp1Retracted : BOOL;
    bDp2Retracted : BOOL;
    abChainSlack : ARRAY[1..4] OF BOOL;
END_STRUCT
END_TYPE

// ---- DUTs/HMI/ST_VTD_ManualHmiCommand.TcDUT
// HMI -> PLC: commands of the VTD manual test screen VTD_ManualTest (TEST ONLY).
// Read by FB_VTD_ManualControl. The PLC writes back:
//  - bEnable       reset to FALSE when the enable is dropped (no automatic restart)
//  - eModeRequest  set to the active mode after every evaluation
//  - iSpeedPercent limited to 0..100
TYPE ST_VTD_ManualHmiCommand :
STRUCT
    bEnable : BOOL;              // Toggle - drive enable request
    bJogPositive : BOOL;         // Tap, hold-to-run - jog +, modes 100/101
    bJogNegative : BOOL;         // Tap, hold-to-run - jog -, modes 100/101
    bRunPositive : BOOL;         // Tap - run in positive direction, mode 200 (latched in the PLC)
    bRunNegative : BOOL;         // Tap - run in negative direction, mode 200 (latched in the PLC)
    bStart : BOOL;               // Tap - start, modes 300/400/401 (latched in the PLC)
    bStop : BOOL;                // Tap - normal stop with the PO 4 deceleration
    bSoftwareStop : BOOL;        // Tap - SOFTWARE STOP, not a safety function (latched in the PLC)
    bReset : BOOL;               // Tap - clears the software stop and resets drive faults (PO 1.8)

    eModeRequest : E_SEW_MovikitMode := E_SEW_MovikitMode.JogSpeedControlled; // Written by the mode buttons
    iSpeedPercent : INT := 10;   // Speed in % of stManualSettings.iMaxSpeed (0..100)
    diTargetPosition : DINT;     // User units. Mode 400: absolute target, mode 401: relative distance
END_STRUCT
END_TYPE

// ---- DUTs/HMI/ST_VTD_ManualHmiStatus.TcDUT
// PLC -> HMI: status of the VTD manual test screen VTD_ManualTest (TEST ONLY).
// Written by FB_VTD_ManualControl, copied to GVL_HMI_VTD.stManualStatus by MAIN.
TYPE ST_VTD_ManualHmiStatus :
STRUCT
    // Drive (decoded PI 1..8)
    stDrive : ST_SEW_MovikitStatus;
    udiErrorId : UDINT;              // FB_SEW_Drive error id: PI 3 (fault * 256 + subfault) or communication error
    sActualModeName : STRING(40);    // PI 6 as text

    // Operating mode (PO 6)
    eModeActive : E_SEW_MovikitMode;
    sModeActiveName : STRING(40);
    bModeJogPosition : BOOL;         // 100 selected
    bModeJogSpeed : BOOL;            // 101 selected
    bModeSpeed : BOOL;               // 200 selected
    bModeReferencing : BOOL;         // 300 selected
    bModePositionAbsolute : BOOL;    // 400 selected
    bModePositionRelative : BOOL;    // 401 selected
    bModeChangeAllowed : BOOL;       // Standstill and no motion command

    // Command state
    bEnableActive : BOOL;            // Enable sent to the drive (PO 1.0 + PO 1.1)
    bSoftwareStopActive : BOOL;      // Software stop latched, RESET required
    bRawWriteActive : BOOL;          // Raw write of the process data test screen owns the drive
    bSettingsValid : BOOL;           // Max speed, acceleration, deceleration and jog time > 0
    bJogAvailable : BOOL;            // JOG buttons usable
    bRunAvailable : BOOL;            // RUN +/- buttons usable
    bStartAvailable : BOOL;          // START button usable
    bJogPositiveActive : BOOL;       // PO 1.4 requested
    bJogNegativeActive : BOOL;       // PO 1.5 requested
    bJogTimeout : BOOL;              // Jog max time reached, release the button
    bRunPositiveActive : BOOL;
    bRunNegativeActive : BOOL;
    bStartActive : BOOL;             // PO 1.7 requested in modes 300/400/401
    bFaultResetActive : BOOL;        // PO 1.8 pulse running

    // Setpoints sent to the drive
    iSpeedSetpoint : INT;            // PO 2 user units (signed in mode 200, 0 while not enabled)
    diTargetPositionSent : DINT;     // PO 7/8 user units

    // Operator message
    sMessage : STRING(80);
    bMessageAlarm : BOOL;            // TRUE = stop/fault (red), FALSE = information
END_STRUCT
END_TYPE

// ---- DUTs/HMI/ST_VTD_ManualSettings.TcDUT
// Settings of the VTD manual test screen (TEST ONLY). Kept in
// GVL_HMI_VTD.stManualSettings (PERSISTENT) and editable on the screen.
// Speed and ramps are MOVISUITE user units (PO 2..4); the scaling of the VTD is
// not confirmed yet - check the user units in MOVISUITE before entering values.
// 0 = not configured: no motion is accepted until all three values are > 0.
// The application limits configured in MOVISUITE still limit the drive.
TYPE ST_VTD_ManualSettings :
STRUCT
    iMaxSpeed : INT;             // Speed at 100 % on the screen, PO 2 user units (> 0)
    uiAcceleration : UINT;       // PO 3 user units (> 0)
    uiDeceleration : UINT;       // PO 4 user units (> 0)
    tJogMaxTime : TIME := T#30S; // Max continuous jog; the button must be released afterwards
END_STRUCT
END_TYPE

// ---- DUTs/HMI/ST_VTD_PdHmiCommand.TcDUT
// HMI -> PLC: VTD MOVIPRO process data test commands (TEST ONLY screen).
TYPE ST_VTD_PdHmiCommand :
STRUCT
    bTestWriteEnable : BOOL;                  // TEST ONLY - allow PO 2..8
    bTestAllowControlWord : BOOL;             // TEST ONLY - additionally allow PO 1
    aTestProcessOutput : ARRAY[1..8] OF UINT; // TEST ONLY - raw PO 1..8 values
END_STRUCT
END_TYPE

// ---- DUTs/HMI/ST_VTD_PdHmiStatus.TcDUT
// PLC -> HMI: VTD MOVIPRO process data test status (TEST ONLY screen).
// All values are raw; units and bit meanings are pending SEW.
TYPE ST_VTD_PdHmiStatus :
STRUCT
    // Communication
    bCommunicationOk : BOOL;
    bWcStateError : BOOL;
    uiEcState : UINT;                       // 8 = OP
    udiInputChangeCount : UDINT;

    // Process inputs (drive -> PLC)
    aProcessInputRaw : ARRAY[1..8] OF UINT; // PI 1..8
    wStatusWord : WORD;                     // PI 1
    iActualSpeedRaw : INT;                  // PI 2
    wFaultCode : WORD;                      // PI 3
    iTorqueRaw : INT;                       // PI 4
    wDigitalInputs : WORD;                  // PI 5
    uiActualApplicationMode : UINT;         // PI 6
    sActualModeName : STRING(40);           // PI 6 as text (FC_SEW_MovikitModeName)
    diActualPositionRaw : DINT;             // PI 7 (high) + PI 8 (low), user units pending SEW

    // TEST ONLY write
    bTestWriteActive : BOOL;
    bTestWriteExpired : BOOL;
    tTestWriteElapsed : TIME;
    aProcessOutputSent : ARRAY[1..8] OF UINT; // PO 1..8 really sent to the drive
END_STRUCT
END_TYPE

// ---- DUTs/Level_Keys_DUT.TcDUT
TYPE Level_Keys_DUT :
STRUCT
	Level:	ARRAY[1..6] OF BOOL;
END_STRUCT
END_TYPE

// ---- DUTs/Profiling_Station_DUT.TcDUT
TYPE Profiling_Station_DUT :
STRUCT
	Start:  BOOL;
	Ready:  BOOL;
	Running:  Bool;
	Done:  Bool;
	Valid:  Bool;
	OverWidth:  Bool;
	OverHeight:  Bool;
	OverLength:  Bool;
	Error_ID:  Word;
END_STRUCT
END_TYPE

// ---- DUTs/Safety_Stops/Sfts_Control_DUT.TcDUT
TYPE Sfts_Control_DUT :
STRUCT
	Mode:  UINT;
	Error:  BOOL;
	Enabled:  Bool;
	Running:  Bool;
	LP_State:  USInt;
	Motor_Extend:  Bool;
	Motor_Retract:  Bool;
	SM_State:  UInt;
	Instruction:  Sfts_Instruction_DUT;
	Inputs:  Sfts_Inputs_DUT;
END_STRUCT
END_TYPE

// ---- DUTs/Safety_Stops/Sfts_Inputs_DUT.TcDUT
TYPE Sfts_Inputs_DUT :
STRUCT
	DP_Extended:  BOOL;
	DP_Retracted:  Bool;
END_STRUCT
END_TYPE

// ---- DUTs/Safety_Stops/Sfts_Instruction_DUT.TcDUT
TYPE Sfts_Instruction_DUT :
STRUCT
	Mode_Change:  UINT;
	Enable:  BOOL;
	Extend:  Bool;
	Retract:  Bool;
	Manual_Extend:  Bool;
	Manual_Retract:  BOOL;
END_STRUCT
END_TYPE

// ---- DUTs/Safety_Stops/Sfts_Settings_DUT.TcDUT
TYPE Sfts_Settings_DUT :
STRUCT
	ID:  DINT;
	LP_Timeout:  UInt;
END_STRUCT
END_TYPE

// ---- DUTs/SEW/E_SEW_MovikitMode.TcDUT
// MOVIKIT Positioning operating modes (PO 6 setpoint / PI 6 actual).
// Source: SEW manual 33959862, chapter 8.1 "Operating modes".
{attribute 'qualified_only'}
TYPE E_SEW_MovikitMode :
(
    DefaultMode := 0,                    // Enabling or disabling the axes
    JogPositionControlled := 100,        // FCB 20, encoder feedback required
    JogSpeedControlled := 101,           // FCB 05
    Speed := 200,                        // FCB 05
    ReferencingOffsetConfigured := 300,  // FCB 12
    ReferencingOffsetFieldbus := 301,    // FCB 12
    PositioningAbsolute := 400,          // FCB 09
    PositioningRelative := 401,          // FCB 09
    PositioningModuloPositive := 402,    // FCB 09
    PositioningModuloNegative := 403,    // FCB 09
    PositioningModuloShort := 404,       // FCB 09
    TouchprobeAbsoluteDirection := 420,  // FCB 09
    TouchprobeAbsoluteSign := 421,       // FCB 09
    TouchprobeEndlessDirection := 422,   // FCB 09
    TouchprobeEndlessSign := 423,        // FCB 09
    BrakeTest := 700                     // FCB 21
) UINT;
END_TYPE

// ---- DUTs/SEW/ST_SEW_MovikitStatus.TcDUT
// Decoded process input data of a MOVIKIT Positioning drive (Standard 8 PD).
// Source: SEW manual 33959862, chapter 9.5. Written by FB_SEW_Drive.
TYPE ST_SEW_MovikitStatus :
STRUCT
    // Communication
    bEtherCatOk : BOOL;                 // EtherCAT OP and working counter valid
    bHandshakeError : BOOL;             // PI 1.15 did not follow PO 1.15 within the timeout
    bCommunicationOk : BOOL;            // bEtherCatOk AND NOT bHandshakeError

    // PI 1 - Status word
    wStatusWord : WORD;
    bReady : BOOL;                      // PI 1.0
    bStoInactive : BOOL;                // PI 1.1
    bOutputStageEnabled : BOOL;         // PI 1.2
    bBrakeReleased : BOOL;              // PI 1.3
    bMotorTurning : BOOL;               // PI 1.4
    bReferenced : BOOL;                 // PI 1.5
    bRelativePositionApplied : BOOL;    // PI 1.6
    bInPosition : BOOL;                 // PI 1.7
    bError : BOOL;                      // PI 1.8
    bWarning : BOOL;                    // PI 1.9
    bDriveTrain2Active : BOOL;          // PI 1.10
    bSpeedReached : BOOL;               // PI 1.11 setpoint/actual speed comparison
    bSwLimitSwitchesInactive : BOOL;    // PI 1.12
    bStandbyActive : BOOL;              // PI 1.14
    bHandshakeOut : BOOL;               // PI 1.15

    // PI 2..8
    iActualSpeed : INT;                 // PI 2, user units (scaling from MOVISUITE)
    byFaultCode : BYTE;                 // PI 3 high byte (error/warning code)
    bySubfaultCode : BYTE;              // PI 3 low byte (subfault, or active FCB if no error)
    iActualTorque_0p1pct : INT;         // PI 4, 0.1 % of nominal motor torque
    wDigitalInputs : WORD;              // PI 5, DI 00..
    uiActualMode : UINT;                // PI 6, see E_SEW_MovikitMode
    diActualPosition : DINT;            // PI 7 (high) + PI 8 (low), user units
END_STRUCT
END_TYPE

// ---- DUTs/SEW/ST_SEW_ProcessInput5.TcDUT
// Raw process input image of a SEW drive running MOVIKIT Velocity with the
// "5 PD" basic profile, plus the EtherCAT diagnostics of the drive box.
// Source: SEW manual 33959862, chapters 4.2 and 9.5.
TYPE ST_SEW_ProcessInput5 :
STRUCT
    aWord : ARRAY[1..5] OF UINT; // PI 1..5, raw
    bWcStateError : BOOL;        // EtherCAT WcState (TRUE = data invalid)
    uiEcState : UINT;            // EtherCAT InfoData.State (8 = OP)
END_STRUCT
END_TYPE

// ---- DUTs/SEW/ST_SEW_ProcessInput8.TcDUT
// Raw process input image of a SEW drive with the "Standard 8 PD" interface,
// plus the EtherCAT diagnostics of the drive box.
TYPE ST_SEW_ProcessInput8 :
STRUCT
    aWord : ARRAY[1..8] OF UINT; // PI 1..8, raw
    bWcStateError : BOOL;        // EtherCAT WcState (TRUE = data invalid)
    uiEcState : UINT;            // EtherCAT InfoData.State (8 = OP)
END_STRUCT
END_TYPE

// ---- DUTs/SEW/ST_SEW_VelocityScaling.TcDUT
// Scaling and ramps of one SEW MOVIKIT Velocity drive (5 PD), user units from MOVISUITE.
// Same meaning as the SEW fields of Buffer_Cnv_Settings_DUT. 0 = not configured: the motor does not move.
TYPE ST_SEW_VelocityScaling :
STRUCT
	rSewSpeedPerUnit:	REAL;	// PO 2 setpoint [user units] per 1 unit of Cnv_Motor_DUT.Speed
	uiSewAcceleration:	UINT;	// PO 3 acceleration [user units]
	uiSewDeceleration:	UINT;	// PO 4 deceleration [user units]
END_STRUCT
END_TYPE

// ---- DUTs/SEW/ST_SEW_VelocityStatus.TcDUT
// Decoded process input data of a MOVIKIT Velocity drive ("5 PD" profile).
// Source: SEW manual 33959862, chapter 9.5 (only V/P words and bits).
// Written by FB_SEW_VelocityDrive.
TYPE ST_SEW_VelocityStatus :
STRUCT
    // Communication
    bEtherCatOk : BOOL;                 // EtherCAT OP and working counter valid
    bHandshakeError : BOOL;             // PI 1.15 did not follow PO 1.15 within the timeout
    bCommunicationOk : BOOL;            // bEtherCatOk AND NOT bHandshakeError

    // PI 1 - Status word (bits 5, 6, 7 and 12 are MOVIKIT Positioning only)
    wStatusWord : WORD;
    bReady : BOOL;                      // PI 1.0
    bStoInactive : BOOL;                // PI 1.1
    bOutputStageEnabled : BOOL;         // PI 1.2
    bBrakeReleased : BOOL;              // PI 1.3
    bMotorTurning : BOOL;               // PI 1.4
    bError : BOOL;                      // PI 1.8
    bWarning : BOOL;                    // PI 1.9
    bDriveTrain2Active : BOOL;          // PI 1.10
    bSpeedReached : BOOL;               // PI 1.11 setpoint/actual speed comparison
    bStandbyActive : BOOL;              // PI 1.14
    bHandshakeOut : BOOL;               // PI 1.15

    // PI 2..5
    iActualSpeed : INT;                 // PI 2, user units (scaling from MOVISUITE)
    byFaultCode : BYTE;                 // PI 3 high byte (error/warning code)
    bySubfaultCode : BYTE;              // PI 3 low byte (subfault, or active FCB if no error)
    iActualTorque_0p1pct : INT;         // PI 4, 0.1 % of nominal motor torque
    wDigitalInputs : WORD;              // PI 5, DI 00..
END_STRUCT
END_TYPE

// ---- DUTs/Shuttle_Position_UDT.TcDUT
TYPE Shuttle_Position_UDT :
STRUCT
	x: DINT;
	y: DINT;
	Charging: BOOL;
END_STRUCT
END_TYPE

// ---- DUTs/System/E_BarcodeState.TcDUT
{attribute 'qualified_only'}
{attribute 'strict'}
TYPE E_BarcodeState :
(
    Idle := 0,
    Reading := 20,
    Complete := 30
);
END_TYPE

// ---- DUTs/System/ID_Decoded_DUT.TcDUT
TYPE ID_Decoded_DUT :
STRUCT
	Device_Type:  INT;
	Level:  INT;
	VTD:  INT;
END_STRUCT
END_TYPE

// ---- DUTs/System/OrderTable_DUT.TcDUT
TYPE OrderTable_DUT :
STRUCT
	OrderNo:  INT;
	StepNo:  INT;
	PlaceTime:  String[20];
	Device:  String;
	Sequence:  UInt;
	Status:  String[12];
	CompleteTime:  String[20];
	ErrorID:  UInt;
	OPC_Control:  WMS_OPC_UA_DUT;
END_STRUCT
END_TYPE

// ---- DUTs/System/System_DUT.TcDUT
TYPE System_DUT :
STRUCT
	Id:  UINT;
	CancelOrders:  BOOL;
	PauseOrders:  Bool;
	ResumeOrders:  Bool;
	OrderSent:  Bool;
	CurrentOrder:  UInt;
	NextOrder:  UInt;
	OrderTable:  ARRAY[0..99] OF OrderTable_DUT;
	StepTable:  ARRAY[0..20] OF OrderTable_DUT;
	CarParked_Confirm:  Bool;
	Running:  Bool;
	IDLE:  Bool;
	Error:  Bool;
	State:  USInt;
	ResetError:  Bool;
	Ready:  Bool;
	Selected:  Bool;
	Auto_Man:  Bool;
	Paused:  Bool;
// 	Watchdog_TimeOut:  STRUCT;
END_STRUCT
END_TYPE

// ---- DUTs/System/System_Settings_DUT.TcDUT
TYPE System_Settings_DUT :
STRUCT
	VTD_Count:  UINT;
	Level_Count:  UINT;
	Cnv_Count:  UInt;
	Shuttle_Count:  UInt;
	Shuttle_Interlock_Timeout:  UINT;
END_STRUCT
END_TYPE

// ---- DUTs/System/WMS_OPC_UA_DUT.TcDUT
TYPE WMS_OPC_UA_DUT :
STRUCT
	Task_ID:  INT;
	Task_Metadata:  STRING[250];
	Task_Type:  Int;
	Source_Location:  DInt;
	Destination_Location:  DInt;
	Task_Data_Available:  Bool;
	SM_State:  UInt;
	Movement_Ready:  Bool;
	Movement_Request_Complete:  Bool;
	Movement_Request_Complete_Ack:  Bool;
	Shuttle_ID:  Int;
	Shuttle_Loaded:  Bool;
	Pallet_Type:  BYTE;
	Pallet_Alignment:  BYTE;
	SM_State_Maestro:  UInt;
	Pallet_Weight:  INT;
END_STRUCT
END_TYPE

// ---- DUTs/U_DWORD_REAL1.TcDUT
TYPE U_DWORD_REAL1 :
UNION
	dw : DWORD;
    out  : REAL;
END_UNION
END_TYPE

// ---- DUTs/VTD/VTD_Control_DUT.TcDUT
TYPE VTD_Control_DUT :
STRUCT
	Mode:	UINT;
	Error:	BOOL;
	Warning:	UINT;
	Enabled:	BOOL;
	Stopped:	BOOL;
	Running:	BOOL;
	Done:	BOOL;
	Current_Task_Type:	UINT;
	Current_Task_ID:	UINT;
	AbsoluteEnc:	REAL;
	LinearEnc:	REAL;
	Current_Level:	UINT;
	Docked:	BOOL;
	LP_State:	UINT;
	DP_Extended:	BOOL;
	Pallet_Loaded:	UINT;
	Shuttle_Loaded:	UINT;
	SM_State:	UINT;
	Motor_UP:	BOOL;
	Motor_Down:	BOOL;
	Motor_Speed:	UINT;
	VFD_Error:	UINT;
	LE_Error:	UINT;
	AE_Error:	UINT;
	Encoder_Delta:	INT;
	Instruction:	VTD_Instruction_DUT;
	Shuttle_Interlock:	VTD_Shuttle_Interlock_DUT;
	Inputs:	VTD_Inputs_DUT;
	Outputs:	VTD_Outputs_DUT;
	Motor:	VTD_Motor_DUT;
	VTD_Errors:	VTD_Errors_DUT;
END_STRUCT
END_TYPE

// ---- DUTs/VTD/VTD_Errors_DUT.TcDUT
TYPE VTD_Errors_DUT :
STRUCT
	Error_Word_1:	UINT;
	Error_Word_2:	UINT;
	Error_Word_3:	UINT;
	Error_Word_4:	UINT;
	Error_Word_5:	UINT;
END_STRUCT
END_TYPE

// ---- DUTs/VTD/VTD_Inputs_DUT.TcDUT
TYPE VTD_Inputs_DUT :
STRUCT
	Upper_Overtravel:  BOOL;
	Upper_limit:  BOOL;
	Ultimate_SlowDown:  Bool;
	Ultimate_Creep:  Bool;
	Lower_Limit:  Bool;
	Lower_Overtravel:  Bool;
	Level_Detect1:  Bool;
	Level_Detect2:  BOOL;
	DP1_Extended:  BOOL;
	DP2_Extended:  BOOL;
	DP1_Retracted:  BOOL;
	DP2_Retracted:  Bool;
	Chain_Slack_1:  Bool;
	Chain_Slack_2:  Bool;
	Chain_Slack_3:  Bool;
	Chain_Slack_4:  Bool;
	PushToEnter:  Bool;
	PushToExit:  Bool;
	Barcode_1:  STRING;
	Barcode_2:  STRING;
	LE_Status:  UInt;
	LE_Position:  DInt;
	LE_Speed:  Int;
	LE_Warnings:  Int;
	LE_Quality_Decoded_Codes:  Byte;
	LE_Quality_Value:  Byte;
	AE_Status_1:  UInt;
	AE_Status_2:  UInt;
	AE_Position_1:  DInt;
	AE_Position_2:  DInt;
	AE_Speed:  Int;
	VFD_Status:  Word;
	VFD_Speed_Actual:  Word;
	VFD_ActualCurrent:  Int;
	VFD_ActualTorque:  INT;
END_STRUCT
END_TYPE

// ---- DUTs/VTD/VTD_Instruction_DUT.TcDUT
TYPE VTD_Instruction_DUT :
STRUCT
	Mode_Change:  UINT;
	Stop:  BOOL;
	Enable:  Bool;
	Execulte:  Bool;
	Reset:  Bool;
	Pallet_Type:  UInt;
	Task_ID:  UInt;
	Task_Metadata:  String;
	Move_To_Level:  UInt;
	Manual_Up:  Bool;
	Manual_Down:  Bool;
	Manual_LP_Retract:  Bool;
	Manual_LP_Extend:  Bool;
	Start_Teach:  BOOL;
END_STRUCT
END_TYPE

// ---- DUTs/VTD/VTD_Levels_DUT.TcDUT
TYPE VTD_Levels_DUT :
STRUCT
	Levels_LE:	ARRAY[1..8] OF REAL;
END_STRUCT
END_TYPE

// ---- DUTs/VTD/VTD_Motor_DUT.TcDUT
// VTD drive: SEW MOVIPRO with MOVIKIT Positioning Drive, "Standard 8 PD".
// Raw process data is filled by FC Inputs and sent by FC Outputs.
// VTD_FB (via FB_SEW_Drive) writes aProcessOutput and stStatus.
TYPE VTD_Motor_DUT :
STRUCT
	stProcessInput:  ST_SEW_ProcessInput8;  // PI 1..8 + EtherCAT diagnostics, written by Inputs
	aProcessOutput:  ARRAY[1..8] OF UINT;   // PO 1..8 raw, read by Outputs
	stStatus:  ST_SEW_MovikitStatus;        // Decoded drive status, written by VTD_FB
END_STRUCT
END_TYPE

// ---- DUTs/VTD/VTD_Outputs_DUT.TcDUT
TYPE VTD_Outputs_DUT :
STRUCT
	LP1_Retract:  BOOL;
	LP1_Extend:  BOOL;
	LP2_Retract:  Bool;
	LP2_Extend:  Bool;
	AE_Control_Word_1:  WORD;
	AE_Control_Word_2:  WORD;
END_STRUCT
END_TYPE

// ---- DUTs/VTD/VTD_Settings_DUT.TcDUT
TYPE VTD_Settings_DUT :
STRUCT
	ID:  UINT;
	Lowest_Level:  UINT;
	Highest_Level:  UInt;
	VTD_Max_Heigh:  UInt;
	VTD_Min_Height:  UInt;
	VTD_Level_Granularity:  Int;
	Dft_Level_Offset_LE:  Int;
	Dft_Level_Offset_AE:  Int;
	Teach_Speed:  UInt;
	Creep_Speed:  UInt;
	Slow_Speed:  UInt;
	Slow_Calib_Speed:  UInt;
	Loaded_Speed:  UInt;
	Shuttle_Speed:  UInt;
	Pallet_Speed:  UInt;
	Empty_Speed:  UInt;
	Dock_speed:  UInt;
	Manual_Speed:  UInt;
	Slowdown_Count_LE:  UInt;
	Creep_Count_LE:  UInt;
	Slowdown_Count_AE:  UInt;
	Creep_Count_AE:  UInt;
	Encoder_Delta_W1:  Real;
	Encoder_Delta_W2:  Real;
	AE_Ratio:  Real;
	Encoder_Delta_Warning:  Real;
	Encoder_Delta_Error:  Real;
	Transfer_Timeout_Up:  UInt;
	Transfer_Timeout_Down:  UInt;
	Lockpins_Timeout_Extend:  UInt;
	Lockpins_Timeout_Retract:  UInt;
	Level_Detect_Timeout:  UInt;
	Teach_Timeout:  UInt;
	Chain_Slack_Timeout:  UInt;
	Level_Detect_LE:  Real;
	Acc_Range_1:  UInt;
	Acc_Range_2:  UInt;
	Acc_Range_3:  UInt;
	Weight_Range_1:  UInt;
	Weight_Range_2:  UInt;
	Weight_Range_3:  UInt;
	Teach_Values:  VTD_Levels_DUT;
	// SEW MOVIKIT scaling (user units from MOVISUITE). 0 = not configured: the VTD does not move.
	SEW_Speed_At_100pct:  INT;   // PO 2 speed setpoint [user units] for Motor_Speed = 100 %
	SEW_Ramp_At_100pct:  UINT;   // PO 3/PO 4 acceleration/deceleration [user units] for ramp factor = 100 %
END_STRUCT
END_TYPE

// ---- DUTs/VTD/VTD_Shuttle_Interlock_DUT.TcDUT
TYPE VTD_Shuttle_Interlock_DUT :
STRUCT
	Interlock_Complete:  BOOL;
	Interlock_Complete_Ack:  BOOL;
	Ready_To_Interlock:  Bool;
	Interlock_Request:  Bool;
	Shuttle_ID:  UInt;
	Shuttle_Target_Location:  DInt;
	Shuttle_Start_Location:  DInt;
	Shuttle_Loaded:  Bool;
	Shuttle_Interlock_Task_ID:  UInt;
	Shuttle_Interlock_Task_Metadata:  STRING;
END_STRUCT
END_TYPE

// ---- GVLs/Control.TcGVL
{attribute 'qualified_only'}
VAR_GLOBAL
	//DEVICES
	VTD:  VTD_Control_DUT;
	ECnv:  ECnv_Control_DUT;
	LCnv:  ARRAY[1..6] OF Buffer_Cnv_Control_DUT;
	Turn_Table: Turn_Table_Control_DUT;
	TBCnv:  TBCnv_Control_DUT;
	Pop_Up_Cnv: ARRAY[1..2] OF PopUp_Control_DUT;
	Roller_Cnv: ARRAY[1..5] OF Roller_Control_DUT;
	Chain_Cnv: Chain_Control_DUT;
	VTDBarcode_Station:  ARRAY[1..3] OF Barcode_Station_DUT;
	Profiling_Station: ARRAY[1..2] OF Profiling_Station_DUT;
	
	//ORDER TABLES COMMANDS
	VTD_Order_Table:  WMS_OPC_UA_DUT;
	Carousel_Order_Table:  WMS_OPC_UA_DUT;
	
	Shuttles_Position:  ARRAY[1..10] OF Shuttle_Position_UDT;
	
	Gate_Station:  ARRAY[1..2] OF Gate_Station_DUT;
	Charger_Level:  ARRAY[1..6] OF Charger_DUT;
	
	//SAFETY (standard PLC -> TwinSAFE logic)
	SafetyReset: BOOL;	// Safety reset pulse (500 ms) for ErrorAcknowledgement and SEW_Safety_Reset. Written by MAIN, copied to IO_Safety by Outputs.
END_VAR

// ---- GVLs/Errors.TcGVL
{attribute 'qualified_only'}
VAR_GLOBAL
	Error:  BOOL;
	Errors_Profinet_1:  WORD;
	Errors_Profinet_10:  Word;
	Errors_Profinet_11:  Word;
	Errors_Profinet_2:  Word;
	Errors_Profinet_3:  Word;
	Errors_Profinet_4:  Word;
	Errors_Profinet_5:  Word;
	Errors_Profinet_6:  Word;
	Errors_Profinet_7:  Word;
	Errors_Profinet_8:  Word;
	Errors_Profinet_9:  Word;
	Errors_Word_Gates_1:  Word;
	Errors_Word_Gates_2:  Word;
	Errors_Word_LightGuard_1:  Word;
	Errors_Word_Logistex:  Word;
	Errors_Word_Shuttles_1:  Word;
	Errors_Word_Shuttles_2:  Word;
	Erros_Supply_Feedback_1:  Word;
	Erros_Supply_Feedback_2:  Word;
	Erros_Supply_Feedback_3:  Word;
	Erros_Supply_Feedback_4:  Word;
	Erros_Supply_Feedback_5:  Word;
	Erros_Supply_Feedback_6:  Word;
	Erros_Supply_Feedback_7:  Word;
	Erros_Word_OPC_1:  Word;
	Erros_Word_OPC_2:  Word;
	Erros_Word_OPC_3:  Word;
	Erros_Word_OPC_4:  Word;
	Erros_Word_OPC_5:  Word;
	Estop_Error_Word_1:  Word;
	Estop_Error_Word_2:  Word;
	Estop_Error_Word_3:  Word;
	Estop_Error_Word_4:  Word;
	Estop_Error_Word_5:  Word;
	Estop_Error_Word_6:  Word;
	LE_Device_Errors_1:  WORD;
	LE_Device_Errors_2:  WORD;
	LE_Device_Errors_3:  WORD;
	LE_Device_Errors_4:  WORD;
	LE_Device_Errors_5:  WORD;
	LE_Warnings_1:  WORD;
	LE_Warnings_2:  WORD;
	LE_Warnings_3:  WORD;
	LE_Warnings_4:  WORD;
	LE_Warnings_5:  WORD;
	Barcode_Reader_ErrorCode_1:  WORD;
	Barcode_Reader_ErrorCode_1_2:  WORD;
	Barcode_Reader_ErrorCode_2:  WORD;
	Barcode_Reader_ErrorCode_2_2:  WORD;
	Barcode_Reader_ErrorCode_3:  WORD;
	Barcode_Reader_ErrorCode_3_2:  WORD;
	Barcode_Reader_ErrorCode_4:  WORD;
	Barcode_Reader_ErrorCode_4_2:  WORD;
	Barcode_Reader_ErrorCode_5:  WORD;
	Barcode_Reader_ErrorCode_5_2:  WORD;
END_VAR

// ---- GVLs/HMI/CNV_HMI.TcGVL
{attribute 'qualified_only'}
VAR_GLOBAL
	CNV_ID_HMI_Old_1:  DINT;
	CNV_ID_HMI:  DINT;
	CNV_ID_HMI_1:  DINT;
	CNV_ID_HMI_Old:  DInt;
	CNV_In_Out_1:  BOOL;
	CNV_Level_Selected:  UInt;
	CNV_Level_Selected_OLD:  UInt;
	CNV_Motor_Actual_Torque:  Real;
	CNV_Motor_Actual_Torque_1:  REAL;
	CNV_Motor_Current_Actual_HMI:  Real;
	CNV_Motor_Current_Actual_HMI_1:  REAL;
	CNV_Motor_Ready:  Bool;
	CNV_Motor_Ready_1:  BOOL;
	CNV_Motor_Status_HMI:  UInt;
	CNV_Motor_Status_HMI_1:  UINT;
	Cnv_Occupied_HMI:  Bool;
	Cnv_Occupied_HMI_1:  BOOL;
	CNV_System_Selected:  UInt;
	CVTD_CNV2_Selected:  UInt;
	Enable_HMI:  Bool;
	Enable_HMI_1:  Bool;
	Enabled_HMI:  Bool;
	Enabled_HMI_1:  Bool;
	Error_HMI:  Bool;
	Error_HMI_1:  Bool;
	HMI_Light_Guard_Bypass:  Bool;
	Light_Guard_Bypass_1:  Bool;
	Light_Guard_Bypass_2:  Bool;
	Manual_Bwd_HMI:  Bool;
	Manual_Bwd_HMI_1:  Bool;
	Manual_Fwd_HMI:  Bool;
	Manual_Fwd_HMI_1:  Bool;
	Manual_Sfty_Stopper_Down_1:  Bool;
	Manual_Sfty_Stopper_Up_1:  Bool;
	Mode_Change_HMI:  UInt;
	Mode_Change_HMI_1:  UInt;
	Mode_HMI:  UInt;
	Mode_HMI_1:  UInt;
	Motor_Direction_HMI:  UInt;
	Motor_Direction_HMI_1:  UInt;
	Motor_Speed_Actual_HMI:  UInt;
	Motor_Speed_Actual_HMI_1:  UInt;
	Motor_Speed_Requested_HMI:  UInt;
	Motor_Speed_Requested_HMI_1:  UInt;
	Ready_For_Task_HMI:  Bool;
	Ready_For_Task_HMI_1:  Bool;
	Reset_HMI:  Bool;
	Reset_HMI_1:  Bool;
	Running_HMI:  Bool;
	Running_HMI_1:  Bool;
	SM_State_HMI:  UInt;
	SM_State_HMI_1:  UInt;
	Start_Transfer_HMI:  Bool;
	Start_Transfer_HMI_1:  Bool;
	Stop_HMI:  Bool;
	Stopped_HMI:  Bool;
	Stopped_HMI_1:  Bool;
	Transfer_From_ID_HMI:  DInt;
	Transfer_From_ID_HMI_1:  DInt;
	Transfer_To_ID_HMI:  DInt;
	Transfer_To_ID_HMI_1:  DInt;
	UpDown_1:  UInt;
	Warning_HMI:  UInt;
	Warning_HMI_1:  UINT;
END_VAR

// ---- GVLs/HMI/CNV_HMI_IO.TcGVL
{attribute 'qualified_only'}
VAR_GLOBAL
	HMI_CNV_SftyPinDown_1:  BOOL;
	HMI_CNV_SftyPinUp_1:  BOOL;
	HMI_Light_Guard:  Bool;
	HMI_CNV_Forward_1:  Bool;
	HMI_CNV_Backward:  Bool;
	HMI_CNV_Forward:  Bool;
	HMI_CNV_Backward_1:  Bool;
END_VAR

// ---- GVLs/HMI/GVL_HMI_Carousel.TcGVL
// HMI interface of the screen Carrousel.
// Device index: 1..2 = PopUp 1..2, 3..7 = Roller 1..5, 8 = Chain, 9 = Turntable.
// TODO: FC_CarouselHmiUpdate once the carousel DUTs / FBs exist. Until then all values stay 0/FALSE.
{attribute 'qualified_only'}
VAR_GLOBAL
    uiSelected : UINT;                                   // HMI -> PLC: 1..9, see above
    astDevice : ARRAY[1..9] OF ST_HMI_ConveyorStatus;    // PLC -> HMI
    stSelected : ST_HMI_ConveyorStatus;                  // PLC -> HMI: copy of the selected device
    stCommand : ST_HMI_ConveyorCommand;                  // HMI -> PLC: commands for the selected device
END_VAR

// ---- GVLs/HMI/GVL_HMI_CNV.TcGVL
// HMI interface of the screen CNV (extractor + buffer conveyors L1..L6).
// The visualization uses only these variables.
// TODO: FC_CnvHmiUpdate (status from Control.ECnv / Control.LCnv, commands to the selected conveyor)
// once the Control refactor compiles. Until then all values stay 0/FALSE.
{attribute 'qualified_only'}
VAR_GLOBAL
    uiSelected : UINT;                                   // HMI -> PLC: 0 = extractor, 1..6 = buffer level
    astConveyor : ARRAY[0..6] OF ST_HMI_ConveyorStatus;  // PLC -> HMI: 0 = extractor, 1..6 = buffer L1..L6
    stSelected : ST_HMI_ConveyorStatus;                  // PLC -> HMI: copy of the selected conveyor
    stCommand : ST_HMI_ConveyorCommand;                  // HMI -> PLC: commands for the selected conveyor
END_VAR

// ---- GVLs/HMI/GVL_HMI_Gates.TcGVL
// HMI interface of the screen Access_Gates. Requests only; the gate locks are
// controlled by the safety logic (TwinSAFE / Euchner MGB2).
// TODO: FC_GatesHmiUpdate (status from Control.Gate_Station). Until then all values stay 0/FALSE.
{attribute 'qualified_only'}
VAR_GLOBAL
    astGate : ARRAY[1..2] OF ST_HMI_GateStatus;      // PLC -> HMI
    astCommand : ARRAY[1..2] OF ST_HMI_GateCommand;  // HMI -> PLC
END_VAR

// ---- GVLs/HMI/GVL_HMI_System.TcGVL
// HMI interface of the system overview (screen Main). The visualization uses only
// these variables; it must not access Control, IO GVLs or FB instances directly.
// TODO: FC_SystemHmiUpdateStatus fills the status from Control once the Control
// refactor (single VTD, carousel DUTs) compiles. Until then all values stay 0/FALSE.
{attribute 'qualified_only'}
VAR_GLOBAL
    stStatus : ST_HMI_SystemStatus;                    // PLC -> HMI
    stCommand : ST_HMI_SystemCommand;                  // HMI -> PLC
    stVtd : ST_HMI_VtdOverview;                        // PLC -> HMI
    stExtractor : ST_HMI_DeviceSummary;                // PLC -> HMI
    astBuffer : ARRAY[1..6] OF ST_HMI_DeviceSummary;   // PLC -> HMI, buffer levels L1..L6
    astPopUp : ARRAY[1..2] OF ST_HMI_DeviceSummary;    // PLC -> HMI, carousel popups
    astRoller : ARRAY[1..5] OF ST_HMI_DeviceSummary;   // PLC -> HMI, carousel rollers
    stChain : ST_HMI_DeviceSummary;                    // PLC -> HMI, carousel chain transfer
    stTurntable : ST_HMI_DeviceSummary;                // PLC -> HMI
    astGate : ARRAY[1..2] OF ST_HMI_GateSummary;       // PLC -> HMI
END_VAR

// ---- GVLs/HMI/GVL_HMI_VTD.TcGVL
// HMI interface of the VTD. The visualization uses only these variables;
// it must not access IO GVLs or FB instances directly.
{attribute 'qualified_only'}
VAR_GLOBAL
    // Screen "Visualization" - process data test (TEST ONLY)
    stPdStatus : ST_VTD_PdHmiStatus;   // PLC -> HMI, written by FC_VTD_PdHmiUpdateStatus
    stPdCommand : ST_VTD_PdHmiCommand; // HMI -> PLC, read by MAIN (TEST ONLY)

    // Screen "VTD_ManualTest" - manual control (TEST ONLY)
    stManualCommand : ST_VTD_ManualHmiCommand; // HMI -> PLC, read and partly written back by FB_VTD_ManualControl
    stManualStatus : ST_VTD_ManualHmiStatus;   // PLC -> HMI, written by MAIN

    // Screen "VTD" - operation
    stStatus : ST_HMI_VtdStatus;     // PLC -> HMI (TODO: FC_VtdHmiUpdate after the Control refactor)
    stCommand : ST_HMI_VtdCommand;   // HMI -> PLC
END_VAR

VAR_GLOBAL PERSISTENT
    stManualSettings : ST_VTD_ManualSettings;  // HMI <-> PLC, test settings kept over a restart
END_VAR

// ---- GVLs/IO/IO_Cards.TcGVL
{attribute 'qualified_only'}
VAR_GLOBAL
	// Source: INBOUND VTD ELECTRICAL DRAWING_9_17_26.pdf, sheets 24.0-27.0.
	// Local PLC rack cards only. Remote module signals belong in a separate IO_Remote GVL.
	// Channel comments identify physical terminals, not PLC process-image offsets.
	// AT %I* / AT %Q* declarations require individual channel links in TwinCAT XAE.
	// Spare outputs are reserved; do not use them in control logic.

	// DI-01 (EL1809) - card 23.0-1, sheet 24.0.
	// Existing REDUNDANCY_OK_8PS1 name retained; the drawing identifies redundancy module 8RS1.
	REDUNDANCY_OK_8PS1 AT %I* : BOOL; // DI-01 CH01 | Wire 24.01 | 8RS1 redundancy OK
	HANDHELD_HMI_KEY_SWITCH_1_NO AT %I* : BOOL; // DI-01 CH02 | Wire 24.02
	HANDHELD_HMI_KEY_SWITCH_2_NO AT %I* : BOOL; // DI-01 CH03 | Wire 24.03
	HANDHELD_HMI_CONNECTED AT %I* : BOOL; // DI-01 CH04 | Wire 24.04
	LM3_4_FAULT AT %I* : BOOL; // DI-01 CH05 | Wire 24.05
	LM5_6_FAULT AT %I* : BOOL; // DI-01 CH06 | Wire 24.06
	LM7_8_FAULT AT %I* : BOOL; // DI-01 CH07 | Wire 24.07
	LM9_FAULT AT %I* : BOOL; // DI-01 CH08 | Wire 24.08
	LM10_FAULT AT %I* : BOOL; // DI-01 CH09 | Wire 24.09
	LM11_FAULT AT %I* : BOOL; // DI-01 CH10 | Wire 24.10
	LM12_FAULT AT %I* : BOOL; // DI-01 CH11 | Wire 24.11
	LM13_14_FAULT AT %I* : BOOL; // DI-01 CH12 | Wire 24.12
	LM15_FAULT AT %I* : BOOL; // DI-01 CH13 | Wire 24.13
	
	LM16_FAULT AT %I* : BOOL; // DI-01 CH14 | Wire 24.14
	_8PS1_OUT_100 AT %I* : BOOL; // DI-01 CH15 | Wire 24.15
	_8PS1_DC_OK AT %I* : BOOL; // DI-01 CH16 | Wire 24.16

	// DI-02 (EL1809) - card 23.0-2, sheet 25.0.
	BACKUP_SIGNAL_BU AT %I* : BOOL; // DI-02 CH01 | Wire 25.01
	TROUBLE_SIGNAL_TR AT %I* : BOOL; // DI-02 CH02 | Wire 25.02
	BATTERY_LOW_SIGNAL_BL AT %I* : BOOL; // DI-02 CH03 | Wire 25.03
	BATTERY_REPLACEMENT_WB AT %I* : BOOL; // DI-02 CH04 | Wire 25.04
	_8PS2_100 AT %I* : BOOL; // DI-02 CH05 | Wire 25.05
	_8PS2_DC_OK AT %I* : BOOL; // DI-02 CH06 | Wire 25.06
	_8PS3_100 AT %I* : BOOL; // DI-02 CH07 | Wire 25.07
	_8PS3_DC_OK AT %I* : BOOL; // DI-02 CH08 | Wire 25.08
	LM100_FAULT AT %I* : BOOL; // DI-02 CH09 | Wire 25.09
	LM101_FAULT AT %I* : BOOL; // DI-02 CH10 | Wire 25.10
	LM102_FAULT AT %I* : BOOL; // DI-02 CH11 | Wire 25.11
	LM103_FAULT AT %I* : BOOL; // DI-02 CH12 | Wire 25.12
	LM104_FAULT AT %I* : BOOL; // DI-02 CH13 | Wire 25.13
	LM105_FAULT AT %I* : BOOL; // DI-02 CH14 | Wire 25.14
	LM106_FAULT AT %I* : BOOL; // DI-02 CH15 | Wire 25.15
	LM107_FAULT AT %I* : BOOL; // DI-02 CH16 | Wire 25.16

	// DO-01 (EL2809) - card 23.0-3, sheet 26.0.
	LM3_16_SET_RESET AT %Q* : BOOL; // DO-01 CH01 | Wire 26.01 | Relay 26CR1
	_50K50_BEACON_INDICATOR_RED AT %Q* : BOOL; // DO-01 CH02 | Wire 26.02 | Relay 26CR2
	_50K50_BEACON_INDICATOR_YELLOW AT %Q* : BOOL; // DO-01 CH03 | Wire 26.03 | Relay 26CR3
	_50K50_BEACON_INDICATOR_GREEN AT %Q* : BOOL; // DO-01 CH04 | Wire 26.04 | Relay 26CR4
	_50K50_BEACON_BUZZER AT %Q* : BOOL; // DO-01 CH05 | Wire 26.05 | Relay 26CR5
	LM100_107_SET_RESET AT %Q* : BOOL; // DO-01 CH06 | Wire 26.06 | Relay 26CR6
	BYPASS_1_FROM_DIGITAL_PLC_OUTPUT AT %Q* : BOOL; // DO-01 CH07 | Wire 26.07 | Relay 26CR7 | Existing safety-interface signal; no bypass logic added
	BYPASS_2_FROM_DIGITAL_PLC_OUTPUT AT %Q* : BOOL; // DO-01 CH08 | Wire 26.08 | Relay 26CR8 | Existing safety-interface signal; no bypass logic added
	BUZZER AT %Q* : BOOL; // DO-01 CH09 | Wire 26.09 | Relay 26CR9
	DO_01_SPARE_CH10 AT %Q* : BOOL; // DO-01 CH10 | Wire 26.10 | Relay 26CR10 | Spare
	DO_01_SPARE_CH11 AT %Q* : BOOL; // DO-01 CH11 | Wire 26.11 | Relay 26CR11 | Spare
	DO_01_SPARE_CH12 AT %Q* : BOOL; // DO-01 CH12 | Wire 26.12 | Relay 26CR12 | Spare
	DO_01_SPARE_CH13 AT %Q* : BOOL; // DO-01 CH13 | Wire 26.13 | Relay 26CR13 | Spare
	DO_01_SPARE_CH14 AT %Q* : BOOL; // DO-01 CH14 | Wire 26.14 | Relay 26CR14 | Spare
	DO_01_SPARE_CH15 AT %Q* : BOOL; // DO-01 CH15 | Wire 26.15 | Relay 26CR15 | Spare
	DO_01_SPARE_CH16 AT %Q* : BOOL; // DO-01 CH16 | Wire 26.16 | Relay 26CR16 | Spare

	// DO-02 (EL2809) - card 23.0-4, sheet 27.0.
	// UPS control uses CH15/CH16. CH01-CH14 are spare.
	DO_02_SPARE_CH01 AT %Q* : BOOL; // DO-02 CH01 | Wire 27.01 | Relay 27CR1 | Spare
	DO_02_SPARE_CH02 AT %Q* : BOOL; // DO-02 CH02 | Wire 27.02 | Relay 27CR2 | Spare
	DO_02_SPARE_CH03 AT %Q* : BOOL; // DO-02 CH03 | Wire 27.03 | Relay 27CR3 | Spare
	DO_02_SPARE_CH04 AT %Q* : BOOL; // DO-02 CH04 | Wire 27.04 | Relay 27CR4 | Spare
	DO_02_SPARE_CH05 AT %Q* : BOOL; // DO-02 CH05 | Wire 27.05 | Relay 27CR5 | Spare
	DO_02_SPARE_CH06 AT %Q* : BOOL; // DO-02 CH06 | Wire 27.06 | Relay 27CR6 | Spare
	DO_02_SPARE_CH07 AT %Q* : BOOL; // DO-02 CH07 | Wire 27.07 | Relay 27CR7 | Spare
	DO_02_SPARE_CH08 AT %Q* : BOOL; // DO-02 CH08 | Wire 27.08 | Relay 27CR8 | Spare
	DO_02_SPARE_CH09 AT %Q* : BOOL; // DO-02 CH09 | Wire 27.09 | Relay 27CR9 | Spare
	DO_02_SPARE_CH10 AT %Q* : BOOL; // DO-02 CH10 | Drawing labels wire 27.27 and relay 27CR27; verify drawing tag. | Spare
	DO_02_SPARE_CH11 AT %Q* : BOOL; // DO-02 CH11 | Wire 27.11 | Relay 27CR11 | Spare
	DO_02_SPARE_CH12 AT %Q* : BOOL; // DO-02 CH12 | Wire 27.12 | Relay 27CR12 | Spare
	DO_02_SPARE_CH13 AT %Q* : BOOL; // DO-02 CH13 | Wire 27.13 | Relay 27CR13 | Spare
	DO_02_SPARE_CH14 AT %Q* : BOOL; // DO-02 CH14 | Wire 27.14 | Relay 27CR14 | Spare
	_8BPS1_REMOTE_ON_OFF AT %Q* : BOOL; // DO-02 CH15 | Wire 27.15 | Relay 27CR15
	_8BPS1_BACKUP_STOP AT %Q* : BOOL; // DO-02 CH16 | Wire 27.16 | Relay 27CR16

	// Existing safety-related declarations below are preserved for compatibility.
	// These standard PLC BOOLs do not implement a safety function.
	// Their relationship to validated TwinSAFE diagnostics must be reviewed before use.
	// See docs/IO_Cards_Review.md for the complete EL1918/EL2912 drawing inventory.
	//FDI-01 (EL1918) - SAFETY INPUTS 23.0-6
	EMERGENCY_STOP_ON_DOOR_CH1 AT%I*:BOOL;
	EMERGENCY_STOP_ON_DOOR_CH2 AT%I*:BOOL;
	EMERGENCY_STOP_ON_HMI AT%I*:BOOL;
END_VAR

// ---- GVLs/IO/IO_Chargers.TcGVL
{attribute 'qualified_only'}
VAR_GLOBAL
// 	Charger Level 1
	Inputs_1 AT%I*:ARRAY[0..19] OF BYTE;
	Outputs_1 AT%Q*:ARRAY[0..9] OF BYTE;
	
	// 	Charger Level 2
	Inputs_2 AT%I*:ARRAY[0..19] OF BYTE;
	Outputs_2 AT%Q*:ARRAY[0..9] OF BYTE;
	
	// 	Charger Level 3
	Inputs_3 AT%I*:ARRAY[0..19] OF BYTE;
	Outputs_3 AT%Q*:ARRAY[0..9] OF BYTE;
	
	// 	Charger Level 4
	Inputs_4 AT%I*:ARRAY[0..19] OF BYTE;
	Outputs_4 AT%Q*:ARRAY[0..9] OF BYTE;
	
	// 	Charger Level 5
	Inputs_5 AT%I*:ARRAY[0..19] OF BYTE;
	Outputs_5 AT%Q*:ARRAY[0..9] OF BYTE;
	
	// 	Charger Level 6
	Inputs_6 AT%I*:ARRAY[0..19] OF BYTE;
	Outputs_6 AT%Q*:ARRAY[0..9] OF BYTE;
	
	// 	Charger Level 7
	Inputs_7 AT%I*:ARRAY[0..19] OF BYTE;
	Outputs_7 AT%Q*:ARRAY[0..9] OF BYTE;
	
	// 	Charger Level 8
	Inputs_8 AT%I*:ARRAY[0..19] OF BYTE;
	Outputs_8 AT%Q*:ARRAY[0..9] OF BYTE;	
END_VAR

// ---- GVLs/IO/IO_RemoteModules.TcGVL
{attribute 'qualified_only'}
VAR_GLOBAL
    // Source: INBOUND VTD ELECTRICAL DRAWING_9_17_26.pdf (rev D), sheets 43.0-48.6 and 53.0-53.5.
    // EtherCAT P remote I/O boxes and TwinSAFE boxes. Local rack cards are in IO_Cards.
    // Box headers give the TwinCAT box name (SpaceX.tsproj) and the drawing tag. The box-to-tag
    // mapping follows the numbering order (confirmed by the user, 2026-10-21).
    // Channel comments: <drawing tag> CH<nn> | <connector> | <description>.
    //   EPP1008: one input per M12 socket X01-X08 (pin 4).
    //   EPP1809: two inputs per M12 socket, X01-X16 (first channel pin 4, second channel pin 2).
    //   EPP2328: four M12 sockets; channel A = pin 4, channel B = pin 2 (sheet 53.0 pinout).
    // AT %I* / AT %Q* declarations require individual channel links in TwinCAT XAE.
    // Spare and unnamed channels are reserved; do not use them in control logic.
    // EtherCAT diagnostics (WcState / EcState) are not linked yet: link them manually in XAE.

    // ---------------------------------------------------------------- Carousel conveyors, EPP1008-0022
    // Sheets 45.0-45.1 / 46.0: boxes for carousel conveyor popups 1-2 and turntable + roller.
    // All EPP1008 channels are shown as '?????????' in drawing rev D: declared as reserved,
    // rename them when the drawing names the signals.
    // 45RIO4 = ENCODER (EPP5001-0002), turntable SSI encoder, sheet 45.5: not part of this GVL.

    // DI-01 (EPP1008-0022) = 45RIO1 - carousel conveyors area section 3 - sheet 45.2.
    _45RIO1_CH01 AT %I* : BOOL; // 45RIO1 CH01 | X01 | Not named in drawing rev D
    _45RIO1_CH02 AT %I* : BOOL; // 45RIO1 CH02 | X02 | Not named in drawing rev D
    _45RIO1_CH03 AT %I* : BOOL; // 45RIO1 CH03 | X03 | Not named in drawing rev D
    _45RIO1_CH04 AT %I* : BOOL; // 45RIO1 CH04 | X04 | Not named in drawing rev D
    _45RIO1_CH05 AT %I* : BOOL; // 45RIO1 CH05 | X05 | Not named in drawing rev D
    _45RIO1_CH06 AT %I* : BOOL; // 45RIO1 CH06 | X06 | Not named in drawing rev D
    _45RIO1_CH07 AT %I* : BOOL; // 45RIO1 CH07 | X07 | Not named in drawing rev D
    _45RIO1_CH08 AT %I* : BOOL; // 45RIO1 CH08 | X08 | Not named in drawing rev D
    _45RIO1_WcState AT %I* : BOOL; // DI-01 > WcState > WcState (TRUE = data invalid)
    _45RIO1_EcState AT %I* : UINT; // DI-01 > InfoData > State (8 = OP)

    // DI-02 (EPP1008-0022) = 45RIO2 - carousel conveyors area section 3 - sheet 45.3.
    _45RIO2_CH01 AT %I* : BOOL; // 45RIO2 CH01 | X01 | Not named in drawing rev D
    _45RIO2_CH02 AT %I* : BOOL; // 45RIO2 CH02 | X02 | Not named in drawing rev D
    _45RIO2_CH03 AT %I* : BOOL; // 45RIO2 CH03 | X03 | Not named in drawing rev D
    _45RIO2_CH04 AT %I* : BOOL; // 45RIO2 CH04 | X04 | Not named in drawing rev D
    _45RIO2_CH05 AT %I* : BOOL; // 45RIO2 CH05 | X05 | Not named in drawing rev D
    _45RIO2_CH06 AT %I* : BOOL; // 45RIO2 CH06 | X06 | Not named in drawing rev D
    _45RIO2_CH07 AT %I* : BOOL; // 45RIO2 CH07 | X07 | Not named in drawing rev D
    _45RIO2_CH08 AT %I* : BOOL; // 45RIO2 CH08 | X08 | Not named in drawing rev D
    _45RIO2_WcState AT %I* : BOOL; // DI-02 > WcState > WcState (TRUE = data invalid)
    _45RIO2_EcState AT %I* : UINT; // DI-02 > InfoData > State (8 = OP)

    // DI-03 (EPP1008-0022) = 45RIO3 - carousel conveyors area section 3 - sheet 45.4.
    _45RIO3_CH01 AT %I* : BOOL; // 45RIO3 CH01 | X01 | Not named in drawing rev D
    _45RIO3_CH02 AT %I* : BOOL; // 45RIO3 CH02 | X02 | Not named in drawing rev D
    _45RIO3_CH03 AT %I* : BOOL; // 45RIO3 CH03 | X03 | Not named in drawing rev D
    _45RIO3_CH04 AT %I* : BOOL; // 45RIO3 CH04 | X04 | Not named in drawing rev D
    _45RIO3_CH05 AT %I* : BOOL; // 45RIO3 CH05 | X05 | Not named in drawing rev D
    _45RIO3_CH06 AT %I* : BOOL; // 45RIO3 CH06 | X06 | Not named in drawing rev D
    _45RIO3_CH07 AT %I* : BOOL; // 45RIO3 CH07 | X07 | Not named in drawing rev D
    _45RIO3_CH08 AT %I* : BOOL; // 45RIO3 CH08 | X08 | Not named in drawing rev D
    _45RIO3_WcState AT %I* : BOOL; // DI-03 > WcState > WcState (TRUE = data invalid)
    _45RIO3_EcState AT %I* : UINT; // DI-03 > InfoData > State (8 = OP)

    // DI-04 (EPP1008-0022) = 46RIO1 - carousel conveyors area sections 1 & 2 - sheet 46.1.
    _46RIO1_CH01 AT %I* : BOOL; // 46RIO1 CH01 | X01 | Not named in drawing rev D
    _46RIO1_CH02 AT %I* : BOOL; // 46RIO1 CH02 | X02 | Not named in drawing rev D
    _46RIO1_CH03 AT %I* : BOOL; // 46RIO1 CH03 | X03 | Not named in drawing rev D
    _46RIO1_CH04 AT %I* : BOOL; // 46RIO1 CH04 | X04 | Not named in drawing rev D
    _46RIO1_CH05 AT %I* : BOOL; // 46RIO1 CH05 | X05 | Not named in drawing rev D
    _46RIO1_CH06 AT %I* : BOOL; // 46RIO1 CH06 | X06 | Not named in drawing rev D
    _46RIO1_CH07 AT %I* : BOOL; // 46RIO1 CH07 | X07 | Not named in drawing rev D
    _46RIO1_CH08 AT %I* : BOOL; // 46RIO1 CH08 | X08 | Not named in drawing rev D
    _46RIO1_WcState AT %I* : BOOL; // DI-04 > WcState > WcState (TRUE = data invalid)
    _46RIO1_EcState AT %I* : UINT; // DI-04 > InfoData > State (8 = OP)

    // DI-05 (EPP1008-0022) = 46RIO2 - carousel conveyors area sections 1 & 2 - sheet 46.2.
    _46RIO2_CH01 AT %I* : BOOL; // 46RIO2 CH01 | X01 | Not named in drawing rev D
    _46RIO2_CH02 AT %I* : BOOL; // 46RIO2 CH02 | X02 | Not named in drawing rev D
    _46RIO2_CH03 AT %I* : BOOL; // 46RIO2 CH03 | X03 | Not named in drawing rev D
    _46RIO2_CH04 AT %I* : BOOL; // 46RIO2 CH04 | X04 | Not named in drawing rev D
    _46RIO2_CH05 AT %I* : BOOL; // 46RIO2 CH05 | X05 | Not named in drawing rev D
    _46RIO2_CH06 AT %I* : BOOL; // 46RIO2 CH06 | X06 | Not named in drawing rev D
    _46RIO2_CH07 AT %I* : BOOL; // 46RIO2 CH07 | X07 | Not named in drawing rev D
    _46RIO2_CH08 AT %I* : BOOL; // 46RIO2 CH08 | X08 | Not named in drawing rev D
    _46RIO2_WcState AT %I* : BOOL; // DI-05 > WcState > WcState (TRUE = data invalid)
    _46RIO2_EcState AT %I* : UINT; // DI-05 > InfoData > State (8 = OP)

    // DI-06 (EPP1008-0022) = 46RIO3 - carousel conveyors area sections 1 & 2 - sheet 46.3.
    _46RIO3_CH01 AT %I* : BOOL; // 46RIO3 CH01 | X01 | Not named in drawing rev D
    _46RIO3_CH02 AT %I* : BOOL; // 46RIO3 CH02 | X02 | Not named in drawing rev D
    _46RIO3_CH03 AT %I* : BOOL; // 46RIO3 CH03 | X03 | Not named in drawing rev D
    _46RIO3_CH04 AT %I* : BOOL; // 46RIO3 CH04 | X04 | Not named in drawing rev D
    _46RIO3_CH05 AT %I* : BOOL; // 46RIO3 CH05 | X05 | Not named in drawing rev D
    _46RIO3_CH06 AT %I* : BOOL; // 46RIO3 CH06 | X06 | Not named in drawing rev D
    _46RIO3_CH07 AT %I* : BOOL; // 46RIO3 CH07 | X07 | Not named in drawing rev D
    _46RIO3_CH08 AT %I* : BOOL; // 46RIO3 CH08 | X08 | Not named in drawing rev D
    _46RIO3_WcState AT %I* : BOOL; // DI-06 > WcState > WcState (TRUE = data invalid)
    _46RIO3_EcState AT %I* : UINT; // DI-06 > InfoData > State (8 = OP)

    // DI-07 (EPP1008-0022) = 46RIO4 - carousel conveyors area sections 1 & 2 - sheet 46.4.
    _46RIO4_CH01 AT %I* : BOOL; // 46RIO4 CH01 | X01 | Not named in drawing rev D
    _46RIO4_CH02 AT %I* : BOOL; // 46RIO4 CH02 | X02 | Not named in drawing rev D
    _46RIO4_CH03 AT %I* : BOOL; // 46RIO4 CH03 | X03 | Not named in drawing rev D
    _46RIO4_CH04 AT %I* : BOOL; // 46RIO4 CH04 | X04 | Not named in drawing rev D
    _46RIO4_CH05 AT %I* : BOOL; // 46RIO4 CH05 | X05 | Not named in drawing rev D
    _46RIO4_CH06 AT %I* : BOOL; // 46RIO4 CH06 | X06 | Not named in drawing rev D
    _46RIO4_CH07 AT %I* : BOOL; // 46RIO4 CH07 | X07 | Not named in drawing rev D
    _46RIO4_CH08 AT %I* : BOOL; // 46RIO4 CH08 | X08 | Not named in drawing rev D
    _46RIO4_WcState AT %I* : BOOL; // DI-07 > WcState > WcState (TRUE = data invalid)
    _46RIO4_EcState AT %I* : UINT; // DI-07 > InfoData > State (8 = OP)

    // DI-08 (EPP1008-0022) = 46RIO5 - carousel conveyors area sections 1 & 2 - sheet 46.5.
    _46RIO5_CH01 AT %I* : BOOL; // 46RIO5 CH01 | X01 | Not named in drawing rev D
    _46RIO5_CH02 AT %I* : BOOL; // 46RIO5 CH02 | X02 | Not named in drawing rev D
    _46RIO5_CH03 AT %I* : BOOL; // 46RIO5 CH03 | X03 | Not named in drawing rev D
    _46RIO5_CH04 AT %I* : BOOL; // 46RIO5 CH04 | X04 | Not named in drawing rev D
    _46RIO5_CH05 AT %I* : BOOL; // 46RIO5 CH05 | X05 | Not named in drawing rev D
    _46RIO5_CH06 AT %I* : BOOL; // 46RIO5 CH06 | X06 | Not named in drawing rev D
    _46RIO5_CH07 AT %I* : BOOL; // 46RIO5 CH07 | X07 | Not named in drawing rev D
    _46RIO5_CH08 AT %I* : BOOL; // 46RIO5 CH08 | X08 | Not named in drawing rev D
    _46RIO5_WcState AT %I* : BOOL; // DI-08 > WcState > WcState (TRUE = data invalid)
    _46RIO5_EcState AT %I* : UINT; // DI-08 > InfoData > State (8 = OP)

    // DI-09 (EPP1008-0022) = 46RIO6 - carousel conveyors area sections 1 & 2 - sheet 46.6.
    _46RIO6_CH01 AT %I* : BOOL; // 46RIO6 CH01 | X01 | Not named in drawing rev D
    _46RIO6_CH02 AT %I* : BOOL; // 46RIO6 CH02 | X02 | Not named in drawing rev D
    _46RIO6_CH03 AT %I* : BOOL; // 46RIO6 CH03 | X03 | Not named in drawing rev D
    _46RIO6_CH04 AT %I* : BOOL; // 46RIO6 CH04 | X04 | Not named in drawing rev D
    _46RIO6_CH05 AT %I* : BOOL; // 46RIO6 CH05 | X05 | Not named in drawing rev D
    _46RIO6_CH06 AT %I* : BOOL; // 46RIO6 CH06 | X06 | Not named in drawing rev D
    _46RIO6_CH07 AT %I* : BOOL; // 46RIO6 CH07 | X07 | Not named in drawing rev D
    _46RIO6_CH08 AT %I* : BOOL; // 46RIO6 CH08 | X08 | Not named in drawing rev D
    _46RIO6_WcState AT %I* : BOOL; // DI-09 > WcState > WcState (TRUE = data invalid)
    _46RIO6_EcState AT %I* : UINT; // DI-09 > InfoData > State (8 = OP)

    // DI-10 (EPP1008-0022) = 46RIO7 - carousel conveyors area sections 1 & 2 - sheet 46.7.
    _46RIO7_CH01 AT %I* : BOOL; // 46RIO7 CH01 | X01 | Not named in drawing rev D
    _46RIO7_CH02 AT %I* : BOOL; // 46RIO7 CH02 | X02 | Not named in drawing rev D
    _46RIO7_CH03 AT %I* : BOOL; // 46RIO7 CH03 | X03 | Not named in drawing rev D
    _46RIO7_CH04 AT %I* : BOOL; // 46RIO7 CH04 | X04 | Not named in drawing rev D
    _46RIO7_CH05 AT %I* : BOOL; // 46RIO7 CH05 | X05 | Not named in drawing rev D
    _46RIO7_CH06 AT %I* : BOOL; // 46RIO7 CH06 | X06 | Not named in drawing rev D
    _46RIO7_CH07 AT %I* : BOOL; // 46RIO7 CH07 | X07 | Not named in drawing rev D
    _46RIO7_CH08 AT %I* : BOOL; // 46RIO7 CH08 | X08 | Not named in drawing rev D
    _46RIO7_WcState AT %I* : BOOL; // DI-10 > WcState > WcState (TRUE = data invalid)
    _46RIO7_EcState AT %I* : UINT; // DI-10 > InfoData > State (8 = OP)

    // ---------------------------------------------------------------- Docking pins and VTD detection

    // DIO-01 (EPP2328-0002) = 47RIO1 - docking pins - sheet 47.3.
    // Outputs go to the docking pins junction box (separate drawing, see note on sheet 47.3).
    // Two signals per socket through Y-cables 6ES7194-6KA00-0XA0 (legs II / III):
    // confirm the leg-to-channel order at the I/O check.
    LEFT_LOCKING_PINS_EXTENDED AT %I* : BOOL; // 47RIO1 CH01 | M12-1 pin 4 | From left locking pins extended proximity sensors
    RIGHT_LOCKING_PINS_EXTENDED AT %I* : BOOL; // 47RIO1 CH02 | M12-1 pin 2 | From right locking pins extended proximity sensors
    LEFT_LOCKING_PINS_RETRACTED AT %I* : BOOL; // 47RIO1 CH03 | M12-2 pin 4 | From left locking pins retracted proximity sensors
    RIGHT_LOCKING_PINS_RETRACTED AT %I* : BOOL; // 47RIO1 CH04 | M12-2 pin 2 | From right locking pins retracted proximity sensors
    DOCKING_PINS_3KA1 AT %Q* : BOOL; // 47RIO1 CH05 | M12-3 pin 4 | To 3KA1 in docking pins junction box
    DOCKING_PINS_3KA2 AT %Q* : BOOL; // 47RIO1 CH06 | M12-3 pin 2 | To 3KA2 in docking pins junction box
    DOCKING_PINS_3KA3 AT %Q* : BOOL; // 47RIO1 CH07 | M12-4 pin 4 | To 3KA3 in docking pins junction box
    DOCKING_PINS_3KA4 AT %Q* : BOOL; // 47RIO1 CH08 | M12-4 pin 2 | To 3KA4 in docking pins junction box
    _47RIO1_WcState AT %I* : BOOL; // DIO-01 > WcState > WcState (TRUE = data invalid)
    _47RIO1_EcState AT %I* : UINT; // DIO-01 > InfoData > State (8 = OP)

    // DI-11 (EPP1809-0022) = 47RIO2 - VTD level, speed and pallet / shuttle detection - sheet 47.4.
    LEVEL_DETECT_1_SENSOR AT %I* : BOOL; // 47RIO2 CH01 | X01 | Level detect 1 sensor
    LEVEL_DETECT_2_SENSOR AT %I* : BOOL; // 47RIO2 CH02 | X02 | Level detect 2 sensor
    CREEP_SENSOR AT %I* : BOOL; // 47RIO2 CH03 | X03 | Creep sensor
    SLOWDOWN_SENSOR AT %I* : BOOL; // 47RIO2 CH04 | X04 | Slowdown sensor
    _47RIO2_CH05 AT %I* : BOOL; // 47RIO2 CH05 | X05 | Wired, not named in drawing rev D
    _47RIO2_SPARE_CH06 AT %I* : BOOL; // 47RIO2 CH06 | X06 | Spare
    _47RIO2_CH07 AT %I* : BOOL; // 47RIO2 CH07 | X07 | Wired, not named in drawing rev D
    _47RIO2_SPARE_CH08 AT %I* : BOOL; // 47RIO2 CH08 | X08 | Spare
    PALLET_DETECTION_1 AT %I* : BOOL; // 47RIO2 CH09 | X09 | Pallet detection #1
    PALLET_DETECTION_2 AT %I* : BOOL; // 47RIO2 CH10 | X10 | Pallet detection #2
    PALLET_DETECTION_3 AT %I* : BOOL; // 47RIO2 CH11 | X11 | Pallet detection #3
    PALLET_DETECTION_4 AT %I* : BOOL; // 47RIO2 CH12 | X12 | Pallet detection #4
    PALLET_DETECTION_5 AT %I* : BOOL; // 47RIO2 CH13 | X13 | Pallet detection #5
    PALLET_DETECTION_6 AT %I* : BOOL; // 47RIO2 CH14 | X14 | Pallet detection #6
    SHUTTLE_DETECTION_1 AT %I* : BOOL; // 47RIO2 CH15 | X15 | Shuttle detection #1
    SHUTTLE_DETECTION_2 AT %I* : BOOL; // 47RIO2 CH16 | X16 | Shuttle detection #2
    _47RIO2_WcState AT %I* : BOOL; // DI-11 > WcState > WcState (TRUE = data invalid)
    _47RIO2_EcState AT %I* : UINT; // DI-11 > InfoData > State (8 = OP)

    // ---------------------------------------------------------------- Buffer conveyors with stopper, EPP2328-0002
    // Outputs drive the coil of stopper motor relays SR8-BB-06A1 (sheets 53.0-53.5).

    // DIO-02 (EPP2328-0002) = 48RIO1 - conveyor with stopper, level 1 - sheets 48.1 and 53.0.
    BUFFER_L1_SAFETY_STOPPER_UPPER_SENSOR AT %I* : BOOL; // 48RIO1 CH01 | M12-1 pin 4 | Safety stopper upper sensor
    BUFFER_L1_SAFETY_STOPPER_LOWER_SENSOR AT %I* : BOOL; // 48RIO1 CH02 | M12-1 pin 2 | Safety stopper lower sensor
    BUFFER_L1_CONVEYOR_SENSOR_1 AT %I* : BOOL; // 48RIO1 CH03 | M12-2 pin 4 | Buffer conveyor sensor 1
    BUFFER_L1_CONVEYOR_SENSOR_2 AT %I* : BOOL; // 48RIO1 CH04 | M12-2 pin 2 | Buffer conveyor sensor 2
    BUFFER_L1_STOPPER_RELAY_53RR1 AT %Q* : BOOL; // 48RIO1 CH05 | M12-3 pin 4 | 53RR1 coil, stopper motor #1 53M1, sheet 53.0/5A
    _48RIO1_SPARE_CH06 AT %Q* : BOOL; // 48RIO1 CH06 | M12-3 pin 2 | Spare
    BUFFER_L1_STOPPER_RELAY_53RR2 AT %Q* : BOOL; // 48RIO1 CH07 | M12-4 pin 4 | 53RR2 coil, sheet 53.0/7E (relay not detailed in drawing rev D)
    _48RIO1_SPARE_CH08 AT %Q* : BOOL; // 48RIO1 CH08 | M12-4 pin 2 | Spare
    _48RIO1_WcState AT %I* : BOOL; // DIO-02 > WcState > WcState (TRUE = data invalid)
    _48RIO1_EcState AT %I* : UINT; // DIO-02 > InfoData > State (8 = OP)

    // DIO-03 (EPP2328-0002) = 48RIO2 - conveyor with stopper, level 2 - sheets 48.2 and 53.1.
    BUFFER_L2_SAFETY_STOPPER_UPPER_SENSOR AT %I* : BOOL; // 48RIO2 CH01 | M12-1 pin 4 | Safety stopper upper sensor
    BUFFER_L2_SAFETY_STOPPER_LOWER_SENSOR AT %I* : BOOL; // 48RIO2 CH02 | M12-1 pin 2 | Safety stopper lower sensor
    BUFFER_L2_CONVEYOR_SENSOR_1 AT %I* : BOOL; // 48RIO2 CH03 | M12-2 pin 4 | Buffer conveyor sensor 1
    BUFFER_L2_CONVEYOR_SENSOR_2 AT %I* : BOOL; // 48RIO2 CH04 | M12-2 pin 2 | Buffer conveyor sensor 2
    BUFFER_L2_STOPPER_RELAY_53RR3 AT %Q* : BOOL; // 48RIO2 CH05 | M12-3 pin 4 | 53RR3 coil, stopper motor #3 53M3, sheet 53.1/5A
    _48RIO2_SPARE_CH06 AT %Q* : BOOL; // 48RIO2 CH06 | M12-3 pin 2 | Spare
    BUFFER_L2_STOPPER_RELAY_53RR4 AT %Q* : BOOL; // 48RIO2 CH07 | M12-4 pin 4 | 53RR4 coil, sheet 53.1/7E (relay not detailed in drawing rev D)
    _48RIO2_SPARE_CH08 AT %Q* : BOOL; // 48RIO2 CH08 | M12-4 pin 2 | Spare
    _48RIO2_WcState AT %I* : BOOL; // DIO-03 > WcState > WcState (TRUE = data invalid)
    _48RIO2_EcState AT %I* : UINT; // DIO-03 > InfoData > State (8 = OP)

    // DIO-04 (EPP2328-0002) = 48RIO3 - conveyor with stopper, level 3 - sheets 48.3 and 53.2.
    BUFFER_L3_SAFETY_STOPPER_UPPER_SENSOR AT %I* : BOOL; // 48RIO3 CH01 | M12-1 pin 4 | Safety stopper upper sensor
    BUFFER_L3_SAFETY_STOPPER_LOWER_SENSOR AT %I* : BOOL; // 48RIO3 CH02 | M12-1 pin 2 | Safety stopper lower sensor
    BUFFER_L3_CONVEYOR_SENSOR_1 AT %I* : BOOL; // 48RIO3 CH03 | M12-2 pin 4 | Buffer conveyor sensor 1
    BUFFER_L3_CONVEYOR_SENSOR_2 AT %I* : BOOL; // 48RIO3 CH04 | M12-2 pin 2 | Buffer conveyor sensor 2
    BUFFER_L3_STOPPER_RELAY_53RR5 AT %Q* : BOOL; // 48RIO3 CH05 | M12-3 pin 4 | 53RR5 coil, stopper motor #5 53M5, sheet 53.2/5A
    _48RIO3_SPARE_CH06 AT %Q* : BOOL; // 48RIO3 CH06 | M12-3 pin 2 | Spare
    BUFFER_L3_STOPPER_RELAY_53RR6 AT %Q* : BOOL; // 48RIO3 CH07 | M12-4 pin 4 | 53RR6 coil, sheet 53.2/7E (relay not detailed in drawing rev D)
    _48RIO3_SPARE_CH08 AT %Q* : BOOL; // 48RIO3 CH08 | M12-4 pin 2 | Spare
    _48RIO3_WcState AT %I* : BOOL; // DIO-04 > WcState > WcState (TRUE = data invalid)
    _48RIO3_EcState AT %I* : UINT; // DIO-04 > InfoData > State (8 = OP)

    // DIO-05 (EPP2328-0002) = 48RIO4 - conveyor with stopper, level 4 - sheets 48.4 and 53.3.
    BUFFER_L4_SAFETY_STOPPER_UPPER_SENSOR AT %I* : BOOL; // 48RIO4 CH01 | M12-1 pin 4 | Safety stopper upper sensor
    BUFFER_L4_SAFETY_STOPPER_LOWER_SENSOR AT %I* : BOOL; // 48RIO4 CH02 | M12-1 pin 2 | Safety stopper lower sensor
    BUFFER_L4_CONVEYOR_SENSOR_1 AT %I* : BOOL; // 48RIO4 CH03 | M12-2 pin 4 | Buffer conveyor sensor 1
    BUFFER_L4_CONVEYOR_SENSOR_2 AT %I* : BOOL; // 48RIO4 CH04 | M12-2 pin 2 | Buffer conveyor sensor 2
    BUFFER_L4_STOPPER_RELAY_53RR7 AT %Q* : BOOL; // 48RIO4 CH05 | M12-3 pin 4 | 53RR7 coil, stopper motor #7 53M7, sheet 53.3/5A
    _48RIO4_SPARE_CH06 AT %Q* : BOOL; // 48RIO4 CH06 | M12-3 pin 2 | Spare
    BUFFER_L4_STOPPER_RELAY_53RR8 AT %Q* : BOOL; // 48RIO4 CH07 | M12-4 pin 4 | 53RR8 coil, sheet 53.3/7E (relay not detailed in drawing rev D)
    _48RIO4_SPARE_CH08 AT %Q* : BOOL; // 48RIO4 CH08 | M12-4 pin 2 | Spare
    _48RIO4_WcState AT %I* : BOOL; // DIO-05 > WcState > WcState (TRUE = data invalid)
    _48RIO4_EcState AT %I* : UINT; // DIO-05 > InfoData > State (8 = OP)

    // DIO-06 (EPP2328-0002) = 48RIO5 - conveyor with stopper, level 5 - sheets 48.5 and 53.4.
    BUFFER_L5_SAFETY_STOPPER_UPPER_SENSOR AT %I* : BOOL; // 48RIO5 CH01 | M12-1 pin 4 | Safety stopper upper sensor
    BUFFER_L5_SAFETY_STOPPER_LOWER_SENSOR AT %I* : BOOL; // 48RIO5 CH02 | M12-1 pin 2 | Safety stopper lower sensor
    BUFFER_L5_CONVEYOR_SENSOR_1 AT %I* : BOOL; // 48RIO5 CH03 | M12-2 pin 4 | Buffer conveyor sensor 1
    BUFFER_L5_CONVEYOR_SENSOR_2 AT %I* : BOOL; // 48RIO5 CH04 | M12-2 pin 2 | Buffer conveyor sensor 2
    BUFFER_L5_STOPPER_RELAY_53RR9 AT %Q* : BOOL; // 48RIO5 CH05 | M12-3 pin 4 | 53RR9 coil, stopper motor #9 53M9, sheet 53.4/5A
    _48RIO5_SPARE_CH06 AT %Q* : BOOL; // 48RIO5 CH06 | M12-3 pin 2 | Spare
    BUFFER_L5_STOPPER_RELAY_53RR10 AT %Q* : BOOL; // 48RIO5 CH07 | M12-4 pin 4 | 53RR10 coil, sheet 53.4/7E (relay not detailed in drawing rev D)
    _48RIO5_SPARE_CH08 AT %Q* : BOOL; // 48RIO5 CH08 | M12-4 pin 2 | Spare
    _48RIO5_WcState AT %I* : BOOL; // DIO-06 > WcState > WcState (TRUE = data invalid)
    _48RIO5_EcState AT %I* : UINT; // DIO-06 > InfoData > State (8 = OP)

    // DIO-07 (EPP2328-0002) = 48RIO6 - conveyor with stopper, level 6 - sheets 48.6 and 53.5.
    BUFFER_L6_SAFETY_STOPPER_UPPER_SENSOR AT %I* : BOOL; // 48RIO6 CH01 | M12-1 pin 4 | Safety stopper upper sensor
    BUFFER_L6_SAFETY_STOPPER_LOWER_SENSOR AT %I* : BOOL; // 48RIO6 CH02 | M12-1 pin 2 | Safety stopper lower sensor
    BUFFER_L6_CONVEYOR_SENSOR_1 AT %I* : BOOL; // 48RIO6 CH03 | M12-2 pin 4 | Buffer conveyor sensor 1
    BUFFER_L6_CONVEYOR_SENSOR_2 AT %I* : BOOL; // 48RIO6 CH04 | M12-2 pin 2 | Buffer conveyor sensor 2
    BUFFER_L6_STOPPER_RELAY_53RR11 AT %Q* : BOOL; // 48RIO6 CH05 | M12-3 pin 4 | 53RR11 coil, stopper motor #11 53M11, sheet 53.5/5A
    _48RIO6_SPARE_CH06 AT %Q* : BOOL; // 48RIO6 CH06 | M12-3 pin 2 | Spare
    BUFFER_L6_STOPPER_RELAY_53RR12 AT %Q* : BOOL; // 48RIO6 CH07 | M12-4 pin 4 | 53RR12 coil, sheet 53.5/7E (relay not detailed in drawing rev D)
    _48RIO6_SPARE_CH08 AT %Q* : BOOL; // 48RIO6 CH08 | M12-4 pin 2 | Spare
    _48RIO6_WcState AT %I* : BOOL; // DIO-07 > WcState > WcState (TRUE = data invalid)
    _48RIO6_EcState AT %I* : UINT; // DIO-07 > InfoData > State (8 = OP)

    // ---------------------------------------------------------------- TwinSAFE boxes
    // Safe channels travel in the FSoE frame to the TwinSAFE logic. They are NOT standard PLC I/O:
    // the standard PLC gets their state only through TwinSAFE logic outputs (IO_Safety).
    // Only diagnostics and the EP1957 standard (non-safe) data are declared here.

    // FDI-01 (EP1918-0002) = 43SRIO1 - safe inputs - sheets 43.0-43.1.
    //   In1/In2: 43SC1 to overtravel upper (NC).
    //   In3/In4: 43SC2 to overtravel lower (NC).
    //   In5-In8: spare.
    _43SRIO1_WcState AT %I* : BOOL; // FDI-01 > WcState > WcState (TRUE = data invalid)
    _43SRIO1_EcState AT %I* : UINT; // FDI-01 > InfoData > State (8 = OP)

    // FDIO-01 (EP1957-0022) = 43SRIO2 - safe inputs / outputs - sheets 43.2-43.4.
    //   In1/In2: 43LC1 light curtain receiver OSSD1 / OSSD2 (SICK C4C-EV13530B10000), sheet 43.4.
    //   In3/In4: 43LC2 light curtain sender (SICK C4C-SV13530B10000), sheet 43.4.
    //   Other safe inputs and safe outputs 1-4: not used in drawing rev D.
    _43SRIO2_SPARE_STD_OUT1 AT %Q* : BOOL; // FDIO-01 > Outputs > Module 1.Standard Output | Spare (no output used in drawing rev D)
    _43SRIO2_SPARE_STD_OUT2 AT %Q* : BOOL; // FDIO-01 > Outputs > Module 2.Standard Output | Spare (no output used in drawing rev D)
    _43SRIO2_SPARE_STD_OUT3 AT %Q* : BOOL; // FDIO-01 > Outputs > Module 3.Standard Output | Spare (no output used in drawing rev D)
    _43SRIO2_SPARE_STD_OUT4 AT %Q* : BOOL; // FDIO-01 > Outputs > Module 4.Standard Output | Spare (no output used in drawing rev D)
    _43SRIO2_FIELDVOLTAGE_UNDERRANGE AT %I* : BOOL; // FDIO-01 > FIELDVOLTAGE Field Voltage Status > Fieldvoltage Underrange
    _43SRIO2_FIELDVOLTAGE_OVERRANGE AT %I* : BOOL; // FDIO-01 > FIELDVOLTAGE Field Voltage Status > Fieldvoltage Overrange
    _43SRIO2_WcState AT %I* : BOOL; // FDIO-01 > WcState > WcState (TRUE = data invalid)
    _43SRIO2_EcState AT %I* : UINT; // FDIO-01 > InfoData > State (8 = OP)
END_VAR

// ---- GVLs/IO/IO_Safety.TcGVL
//{attribute 'qualified_only'}
VAR_GLOBAL
	ErrorAcknowledgement AT %Q*: BOOL;
	Run AT %Q*: BOOL;
	SEW_Safety_Reset	AT %Q*: BOOL;
END_VAR

// ---- GVLs/IO/IO_VFDs.TcGVL
{attribute 'qualified_only'}
VAR_GLOBAL
	
